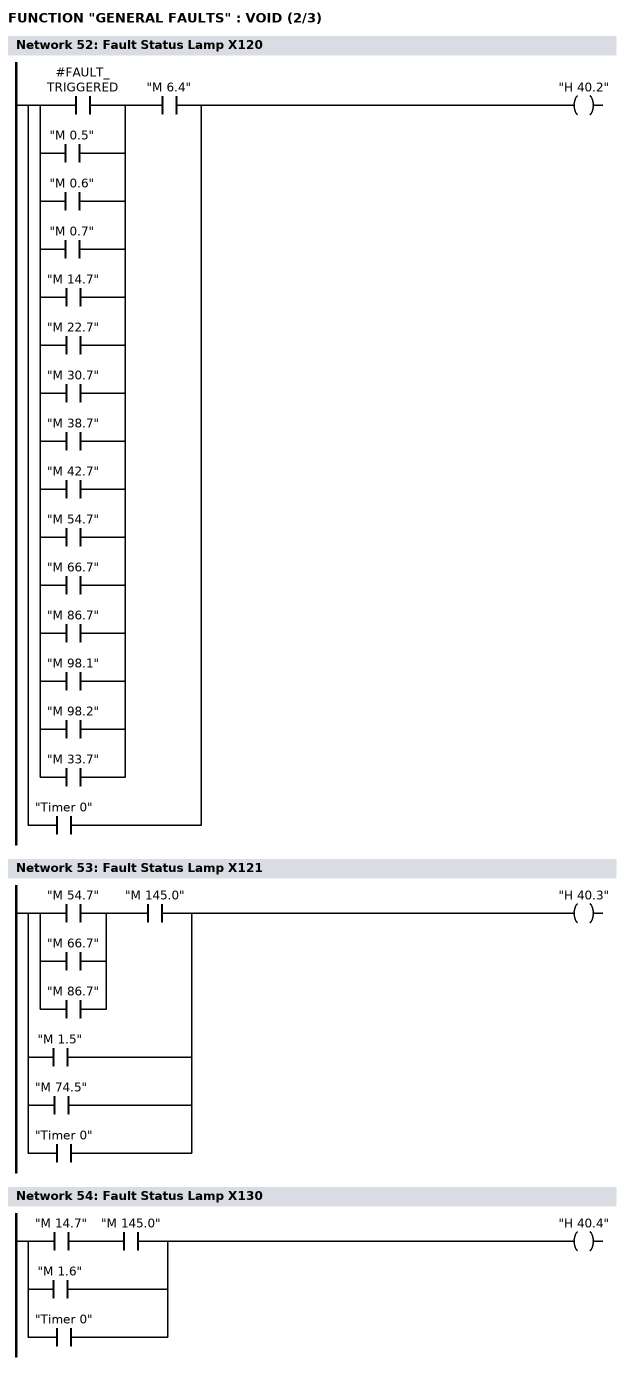

      A(    ;
      O     #FAULT_TRIGGERED;
      O     "M 0.5";
      O     "M 0.6";
      O     "M 0.7";
      O     "M 14.7";
      O     "M 22.7";
      O     "M 30.7";
      O     "M 38.7";
      O     "M 42.7";
      O     "M 54.7";
      O     "M 66.7";
      O     "M 86.7";
      O     "M 98.1";
      O     "M 98.2";
      O     "M 33.7";
      )     ;
      A     "M 6.4";
      O     "Timer 0";
      =     "H 40.2";
NETWORK
TITLE =Fault Status Lamp X121

      A(    ;
      O     "M 54.7";
      O     "M 66.7";
      O     "M 86.7";
      )     ;
      A     "M 145.0";
      O     "M 1.5";
      O     "M 74.5";
      O     "Timer 0";
      =     "H 40.3";
NETWORK
TITLE =Fault Status Lamp X130

      A     "M 14.7";
      A     "M 145.0";
      O     "M 1.6";
      O     "Timer 0";
      =     "H 40.4";
NETWORK
TITLE =Fault Status Lamp X134
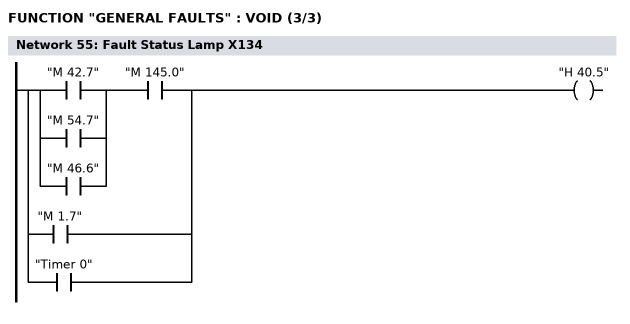

      A(    ;
      O     "M 42.7";
      O     "M 54.7";
      O     "M 46.6";
      )     ;
      A     "M 145.0";
      O     "M 1.7";
      O     "Timer 0";
      =     "H 40.5";
NETWORK
TITLE =Elevator OverTemp

      A     "M 0.6";
      AN    "E 0.3";
      L     W#16#1;
      T     "MB 181";
      BEC   ;
NETWORK
TITLE =Turntable OverTemp

      A     "M 0.6";
      AN    "E 0.4";
      L     W#16#2;
      T     "MB 181";
      BEC   ;
NETWORK
TITLE =Loader OverTemp

      A     "M 0.6";
      AN    "E 0.5";
      L     W#16#3;
      T     "MB 181";
      BEC   ;
NETWORK
TITLE =Conveyor 4 Collator OverTemp

      A     "M 0.6";
      AN    "E 14.0";
      L     W#16#4;
      T     "MB 181";
      BEC   ;
NETWORK
TITLE =Conveyor 6 Delivery OverTemp

      A     "M 0.6";
      AN    "E 14.1";
      L     W#16#5;
      T     "MB 181";
      BEC   ;
NETWORK
TITLE =Pivot Conveyor 10 OverTemp

      A(    ;
      ON    "E 14.2";
      ON    "E 14.3";
      )     ;
      A     "M 0.6";
      O     ;
      A(    ;
      O     "E 14.6";
      O     "E 14.7";
      )     ;
      A     "M 0.6";
      L     W#16#6;
      T     "MB 181";
      BEC   ;
NETWORK
TITLE =OverTemp

      A     "M 0.6";
      A     "E 35.0";
      L     W#16#8;
      T     "MB 181";
      BEC   ;
NETWORK
TITLE =OverTemp

      A     "M 0.6";
      A     "E 35.1";
      L     W#16#9;
      T     "MB 181";
      BEC   ;
NETWORK
TITLE =OverTemp

      A     "M 0.6";
      A     "E 14.6";
      L     W#16#B;
      T     "MB 181";
      BEC   ;
NETWORK
TITLE =OverTemp

      A     "M 0.6";
      A     "E 14.7";
      L     W#16#C;
      T     "MB 181";
      BEC   ;
NETWORK
TITLE =

      A     #FAULT_TRIGGERED;
      A     "M 3.0";
      L     W#16#0;
      T     MB   183;
      BEC   ;
NETWORK
TITLE =

      A     #FAULT_TRIGGERED;
      A     "M 3.1";
      L     W#16#1;
      T     MB   183;
      BEC   ;
NETWORK
TITLE =

      A     #FAULT_TRIGGERED;
      A     "M 3.2";
      L     W#16#2;
      T     MB   183;
      BEC   ;
NETWORK
TITLE =

      A     #FAULT_TRIGGERED;
      A     "M 3.3";
      L     W#16#3;
      T     MB   183;
      BEC   ;
NETWORK
TITLE =

      A     #FAULT_TRIGGERED;
      A     "M 3.4";
      L     W#16#4;
      T     MB   183;
      BEC   ;
NETWORK
TITLE =

      A     #FAULT_TRIGGERED;
      A     "M 3.5";
      L     W#16#5;
      T     MB   183;
      BEC   ;
NETWORK
TITLE =

      A     #FAULT_TRIGGERED;
      A     "M 3.6";
      L     W#16#6;
      T     MB   183;
      BEC   ;
NETWORK
TITLE =

      A     #FAULT_TRIGGERED;
      A     "M 3.7";
      L     W#16#7;
      T     MB   183;
      BEC   ;
NETWORK
TITLE =

      A     #FAULT_TRIGGERED;
      A     "M 4.0";
      L     W#16#8;
      T     MB   182;
      BEC   ;
NETWORK
TITLE =

      A     #FAULT_TRIGGERED;
      A     "M 4.1";
      L     W#16#9;
      T     MB   182;
      BEC   ;
NETWORK
TITLE =

      A     #FAULT_TRIGGERED;
      A     "M 4.2";
      L     W#16#10;
      T     MB   182;
      BEC   ;
NETWORK
TITLE =

      A     #FAULT_TRIGGERED;
      A     "M 4.3";
      L     W#16#11;
      T     MB   182;
      BEC   ;
NETWORK
TITLE =

      A     #FAULT_TRIGGERED;
      A     "M 4.4";
      L     W#16#12;
      T     MB   182;
      BEC   ;
NETWORK
TITLE =

      A     #FAULT_TRIGGERED;
      A     "M 4.5";
      L     W#16#13;
      T     MB   182;
      BEC   ;
NETWORK
TITLE =

      A     #FAULT_TRIGGERED;
      A     "M 4.6";
      L     W#16#14;
      T     MB   182;
      BEC   ;
NETWORK
TITLE =

      L     W#16#0;
      T     "MW 180";
      T     MW   182;
END_FUNCTION

FUNCTION "BLINKER" : VOID
TITLE =Blinker
VERSION : 0.0

BEGIN
NETWORK
TITLE =
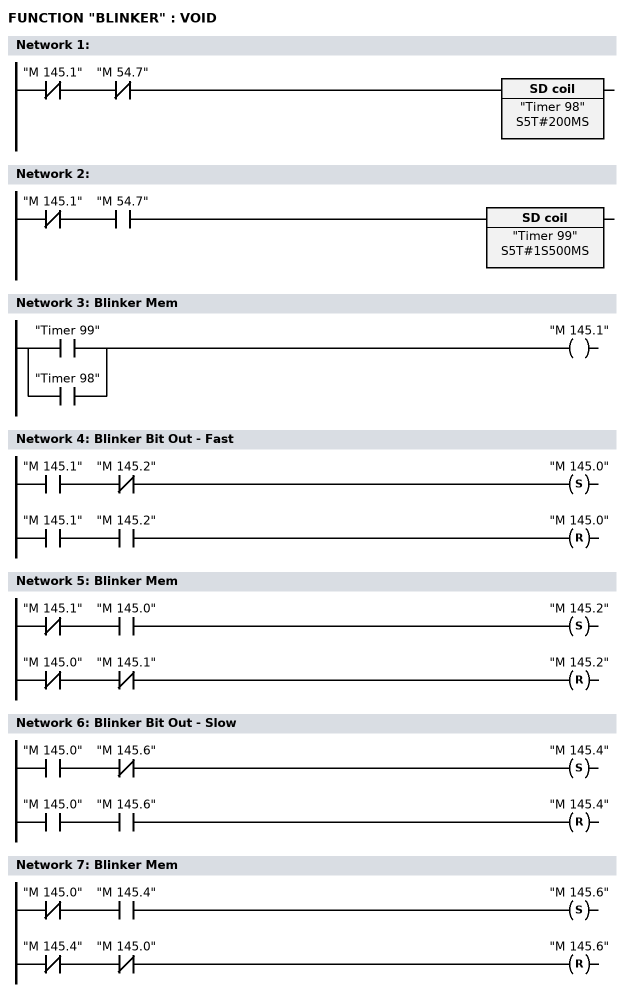

      AN    "M 145.1";
      AN    "M 54.7";
      L     S5T#200MS;
      SD    "Timer 98";
NETWORK
TITLE =

      AN    "M 145.1";
      A     "M 54.7";
      L     S5T#1S500MS;
      SD    "Timer 99";
NETWORK
TITLE =Blinker Mem

      O     "Timer 99";
      O     "Timer 98";
      =     "M 145.1";
NETWORK
TITLE =Blinker Bit Out - Fast

      A     "M 145.1";
      AN    "M 145.2";
      S     "M 145.0";
//;
      A     "M 145.1";
      A     "M 145.2";
      R     "M 145.0";
NETWORK
TITLE =Blinker Mem

      AN    "M 145.1";
      A     "M 145.0";
      S     "M 145.2";
//;
      AN    "M 145.0";
      AN    "M 145.1";
      R     "M 145.2";
NETWORK
TITLE =Blinker Bit Out - Slow

      A     "M 145.0";
      AN    "M 145.6";
      S     "M 145.4";
//;
      A     "M 145.0";
      A     "M 145.6";
      R     "M 145.4";
NETWORK
TITLE =Blinker Mem

      AN    "M 145.0";
      A     "M 145.4";
      S     "M 145.6";
//;
      AN    "M 145.4";
      AN    "M 145.0";
      R     "M 145.6";
END_FUNCTION

FUNCTION "LIGHT CURTAIN - SAFETY" : VOID
TITLE =Conveyors Catways - Access Safety
//Access to Conveyor 1-2-3 & 4 : Crossing Light Curtains Latches / Freezes these
//Conveyors !
//- To Resume Run, CatWay 1 (Conveyors 1-2-3) :  Push Top PB (Catway)
//and Push Lower PB (Main Floor) within 15sec .
//- To Resume Run, CatWay 2 (Conveyors 3-4) :  Push Top PB (Catway) .
//
//If Crossing CatWay 2 Light Curtain while No Conveyors are running, Run will
//resume automatic after 1 sec of free Light Curtain.
//
//Big Red Light will Blink to confirm the Conveyors are disabled / Safe .
VERSION : 0.1

BEGIN
NETWORK
TITLE =Safety Light Curtains -  Trigger 2 - Momentary SF = 1s
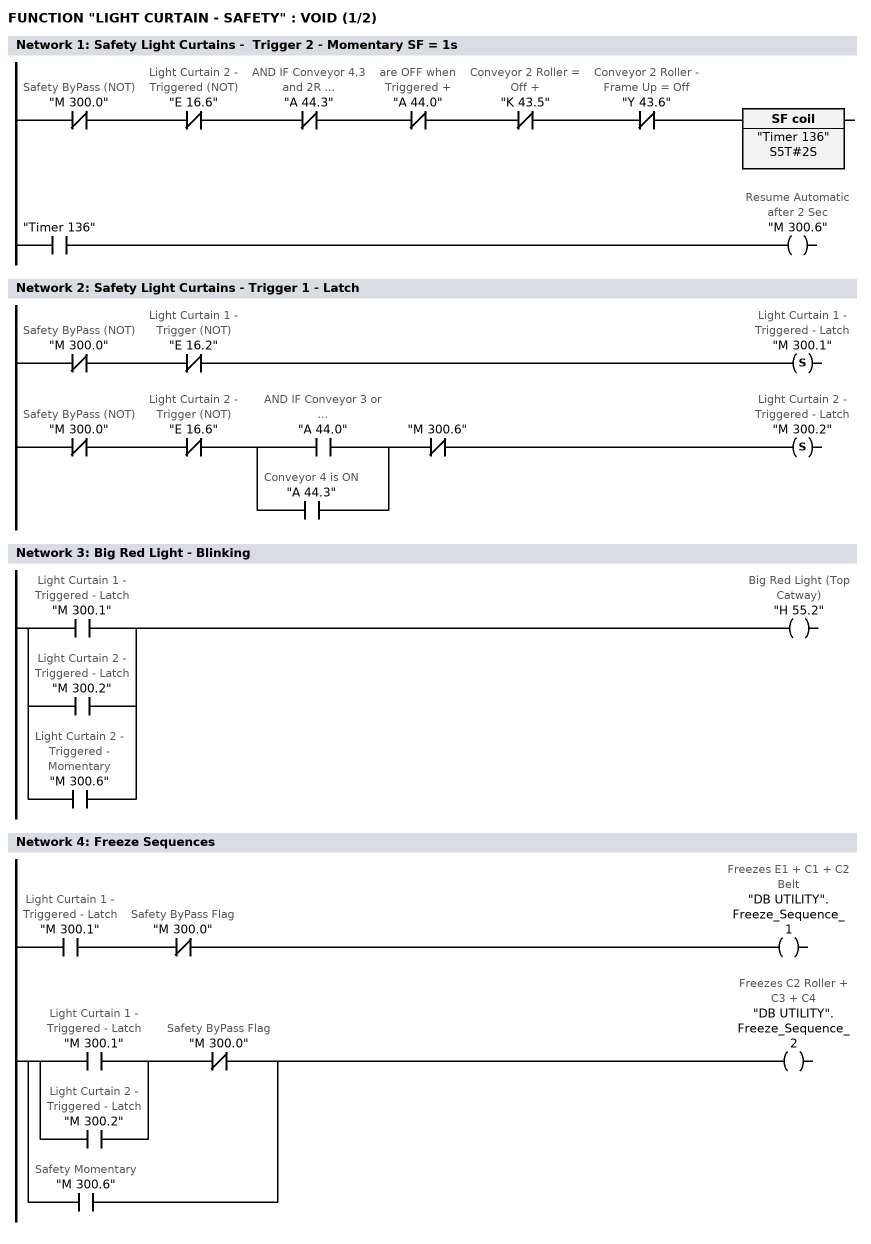

      AN    "M 300.0"; // Safety ByPass (NOT)
      AN    "E 16.6"; // Light Curtain 2 - Triggered (NOT)
      AN    "A 44.3"; // AND IF Conveyor 4,3 and 2R ...
      AN    "A 44.0"; // are OFF when Triggered +
      AN    "K 43.5"; // Conveyor 2 Roller = Off +
      AN    "Y 43.6"; // Conveyor 2 Roller - Frame Up = Off
      L     S5T#2S;
      SF    "Timer 136"; // Debouncer 2s
//;
      A     "Timer 136";
      =     "M 300.6"; // Resume Automatic after 2 Sec

NETWORK
TITLE =Safety Light Curtains - Trigger 1 - Latch

      AN    "M 300.0"; // Safety ByPass (NOT)
      AN    "E 16.2"; // Light Curtain 1 - Trigger (NOT)
      S     "M 300.1"; // Light Curtain 1 - Triggered - Latch
//;
      AN    "M 300.0"; // Safety ByPass (NOT)
      AN    "E 16.6"; // Light Curtain 2 - Trigger (NOT)
      A(    ;
      O     "A 44.0"; // AND IF Conveyor 3 or ...
      O     "A 44.3"; // Conveyor 4 is ON
      )     ;
      AN    "M 300.6";
      S     "M 300.2"; // Light Curtain 2 - Triggered - Latch
NETWORK
TITLE =Big Red Light - Blinking

      A(    ;
      O     "M 300.1"; // Light Curtain 1 - Triggered - Latch
      O     "M 300.2"; // Light Curtain 2 - Triggered - Latch
      O     "M 300.6"; // Light Curtain 2 - Triggered - Momentary
      )     ;
      =     "H 55.2"; // Big Red Light (Top Catway)
NETWORK
TITLE =Freeze Sequences

      A     "M 300.1"; // Light Curtain 1 - Triggered - Latch
      AN    "M 300.0"; // Safety ByPass Flag
      =     "DB UTILITY".Freeze_Sequence_1; //   Freezes E1 + C1 + C2 Belt
//;
      A     "M 300.1"; // Light Curtain 1 - Triggered - Latch
      O     "M 300.2"; // Light Curtain 2 - Triggered - Latch
      AN    "M 300.0"; // Safety ByPass Flag
      O     "M 300.6"; // Safety Momentary
      =     "DB UTILITY".Freeze_Sequence_2; //  Freezes C2 Roller + C3 + C4
NETWORK
TITLE =Safety ByPass - While blocking Curtain, Push Top Button for 5s
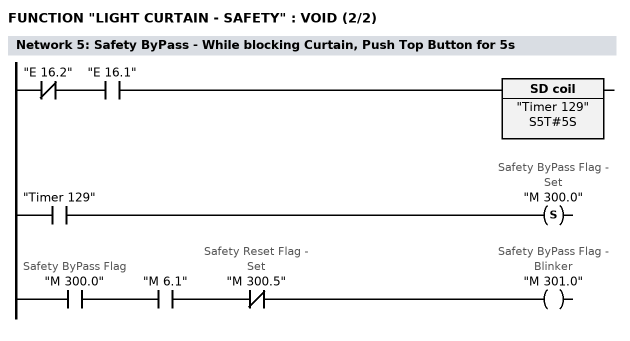

      AN    "E 16.2";
      A     "E 16.1";
      L     S5T#5S;
      SD    "Timer 129";
//;
      A     "Timer 129";
      S     "M 300.0"; // Safety ByPass Flag - Set
//;
      A     "M 300.0"; // Safety ByPass Flag
      A     "M 6.1";
      AN    "M 300.5"; // Safety Reset Flag - Set
      =     "M 301.0"; // Safety ByPass Flag - Blinker

NETWORK
TITLE =TEST REMOTE B+

      R     "A 58.4";

NETWORK
TITLE =PB Led - Control
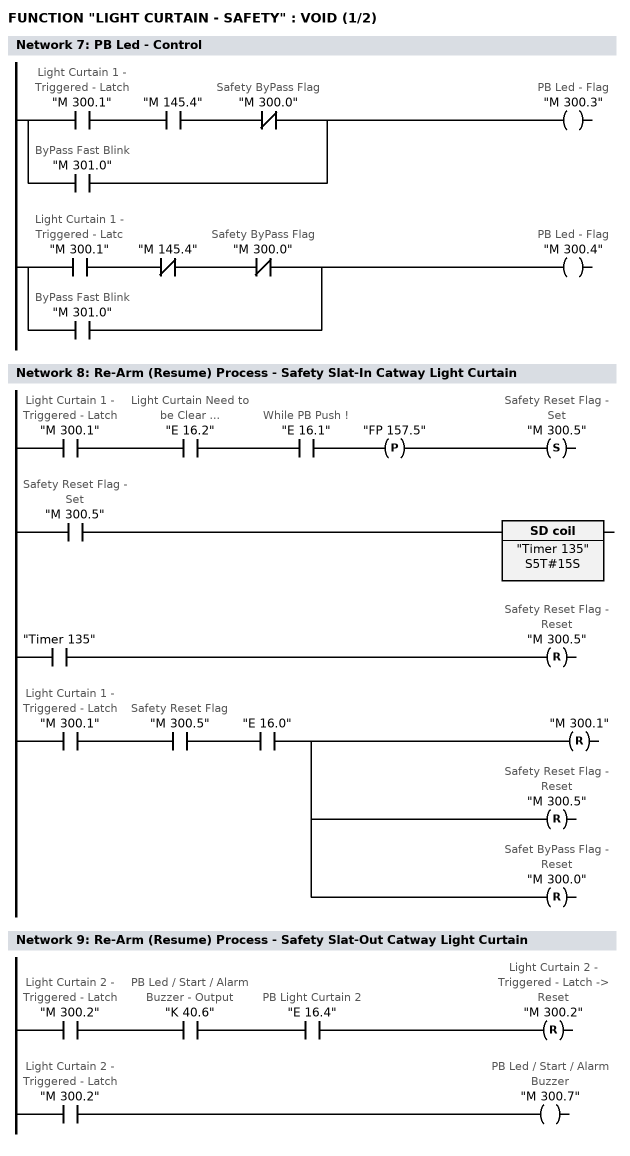

      A     "M 300.1"; // Light Curtain 1 - Triggered - Latch
      A     "M 145.4";
      AN    "M 300.0"; // Safety ByPass Flag
      O     "M 301.0"; // ByPass Fast Blink
      =     "M 300.3"; // PB Led - Flag
//;
      A     "M 300.1"; // Light Curtain 1 - Triggered - Latc
      AN    "M 145.4";
      AN    "M 300.0"; // Safety ByPass Flag
      O     "M 301.0"; // ByPass Fast Blink
      =     "M 300.4"; // PB Led - Flag
NETWORK
TITLE =Re-Arm (Resume) Process - Safety Slat-In Catway Light Curtain

      A     "M 300.1"; // Light Curtain 1 - Triggered - Latch
      A     "E 16.2"; // Light Curtain Need to be Clear ...
      A     "E 16.1"; // While PB Push !
      FP    "FP 157.5";
      S     "M 300.5"; // Safety Reset Flag - Set
//;
      A     "M 300.5"; // Safety Reset Flag - Set
      L     S5T#15S;
      SD    "Timer 135"; // Safety Reset Flag - TimeOut
//;
      A     "Timer 135";
      R     "M 300.5"; // Safety Reset Flag - Reset
//;
      A     "M 300.1"; // Light Curtain 1 - Triggered - Latch
      A     "M 300.5"; // Safety Reset Flag
      A     "E 16.0";
      R     "M 300.1";
      R     "M 300.5"; // Safety Reset Flag - Reset
      R     "M 300.0"; // Safet ByPass Flag - Reset
NETWORK
TITLE =Re-Arm (Resume) Process - Safety Slat-Out Catway Light Curtain

      A     "M 300.2"; // Light Curtain 2 - Triggered - Latch
      A     "K 40.6"; // PB Led / Start / Alarm Buzzer - Output
      A     "E 16.4"; // PB Light Curtain 2
      R     "M 300.2"; // Light Curtain 2 - Triggered - Latch -> Reset
//;
      A     "M 300.2"; // Light Curtain 2 - Triggered - Latch
      =     "M 300.7"; // PB Led / Start / Alarm Buzzer
NETWORK
TITLE =PB Led - Out
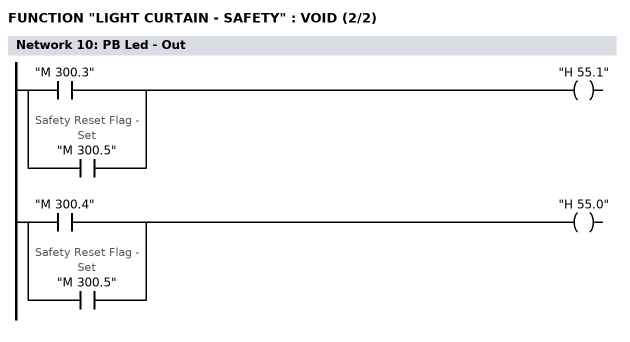

      A     "M 300.3";
      O     "M 300.5"; // Safety Reset Flag - Set
      =     "H 55.1";
//;
      A     "M 300.4";
      O     "M 300.5"; // Safety Reset Flag - Set
      =     "H 55.0";
END_FUNCTION

FUNCTION "CONVEYORS CLEARING" : VOID
TITLE =Conveyors - Clearing Function
//New Order Sequence
NAME : CLEARING
VERSION : 0.0


VAR_TEMP
  EMPTY_11 : BOOL ;	//Empty Conveyor 11
  EMPTY_21 : BOOL ;	//Empty Conveyor 21
  EMPTY_12_22 : BOOL ;	//Empty Conveyor 12 & 22
  EMPTY_13_23 : BOOL ;	//Empty Conveyor 13 & 23
  C10_EMPTY_TEST : BOOL ;
  CLEARING_ABORT : BOOL ;
END_VAR
BEGIN
NETWORK
TITLE =HMI Clearing Call

      A     "M 140.3";
      A     "HMI_DB".CLEARING_SSW_MAIN;
      =     "M 5.2";
//;
      L     8;
      A     "M 10.0";
      =     "HMI_DB".CLEARING_SSW_STATUS;
      JC    CLEA;
      L     0;

CLEA: T     "HMI_DB".CLEARING_FUNCTION;

      A     "M 10.0";
      FN    "FN 155.7";
      R     "HMI_DB".CLEARING_SSW_MAIN;
      R     "M 54.2";
//;
      A     "M 5.2";
      FP    "FP 147.4";
      AN    "B 10.7"; // C11 - Empty
      AN    "B 11.0"; // C12 - Empty
      AN    "B 11.1"; // C13 - Empty
      AN    "B 11.2"; // C13 - Empty
      AN    "B 15.4"; // C21 - Empty
      AN    "B 15.5"; // C22 - Empty
      AN    "B 15.6"; // C23 - Empty
      AN    "B 15.7"; // C23 - Empty
      S     "M 54.2"; // Empty C11...C23
NETWORK
TITLE =New Order Seq - First New Order Packet to Pivot Conveyor 10
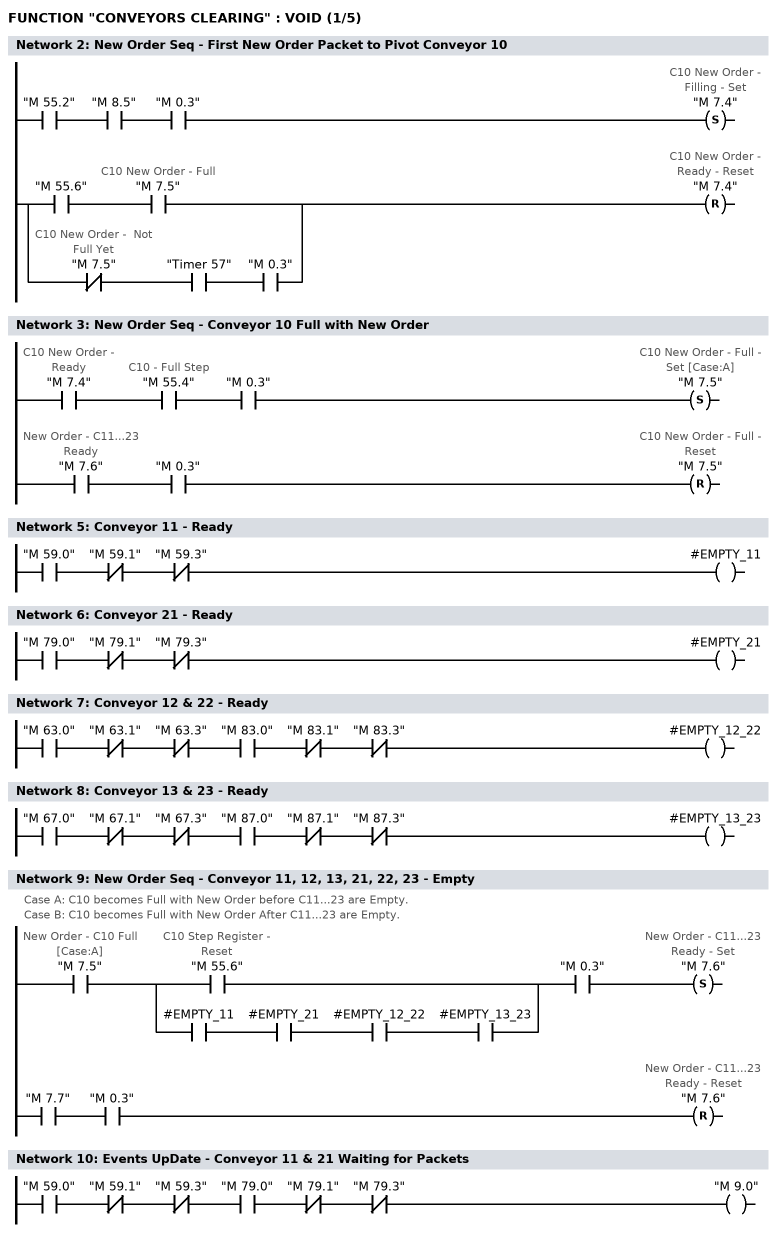

      A     "M 55.2";
      A     "M 8.5";
      A     "M 0.3";
      S     "M 7.4"; // C10 New Order - Filling - Set
//;
      A(    ;
      A     "M 55.6";
      A     "M 7.5"; // C10 New Order - Full
      O     ;
      AN    "M 7.5"; // C10 New Order -  Not Full Yet
      A     "Timer 57";
      A     "M 0.3";
      )     ;
      R     "M 7.4"; // C10 New Order - Ready - Reset
NETWORK
TITLE =New Order Seq - Conveyor 10 Full with New Order

      A     "M 7.4"; // C10 New Order - Ready
      A     "M 55.4"; // C10 - Full Step
      A     "M 0.3";
      S     "M 7.5"; // C10 New Order - Full - Set [Case:A]
//;
      A     "M 7.6"; // New Order - C11...23 Ready
      A     "M 0.3";
      R     "M 7.5"; // C10 New Order - Full - Reset
NETWORK
TITLE =New Order Seq
//New Order Seq - Waiting for the last Order Packets to Run out !


NETWORK
TITLE =Conveyor 11 - Ready

      A     "M 59.0";
      AN    "M 59.1";
      AN    "M 59.3";
      =     #EMPTY_11;
NETWORK
TITLE =Conveyor 21 - Ready

      A     "M 79.0";
      AN    "M 79.1";
      AN    "M 79.3";
      =     #EMPTY_21;
NETWORK
TITLE =Conveyor 12 & 22 - Ready

      A     "M 63.0";
      AN    "M 63.1";
      AN    "M 63.3";
      A     "M 83.0";
      AN    "M 83.1";
      AN    "M 83.3";
      =     #EMPTY_12_22;
NETWORK
TITLE =Conveyor 13 & 23 - Ready

      A     "M 67.0";
      AN    "M 67.1";
      AN    "M 67.3";
      A     "M 87.0";
      AN    "M 87.1";
      AN    "M 87.3";
      =     #EMPTY_13_23;
NETWORK
TITLE =New Order Seq - Conveyor 11, 12, 13, 21, 22, 23 - Empty
//Case A: C10 becomes Full with New Order before C11...23 are Empty.
//Case B: C10 becomes Full with New Order After C11...23 are Empty.
      A     "M 7.5"; // New Order - C10 Full [Case:A]
      A(    ;
      A     "M 55.6"; // C10 Step Register - Reset
      O     ;
      A     #EMPTY_11;
      A     #EMPTY_21;
      A     #EMPTY_12_22;
      A     #EMPTY_13_23;
      )     ;
      A     "M 0.3";
      S     "M 7.6"; // New Order - C11...23 Ready - Set
//;
      A     "M 7.7";
      A     "M 0.3";
      R     "M 7.6"; // New Order - C11...23 Ready - Reset
NETWORK
TITLE =Events UpDate - Conveyor 11 & 21 Waiting for Packets

      A     "M 59.0";
      AN    "M 59.1";
      AN    "M 59.3";
      A     "M 79.0";
      AN    "M 79.1";
      AN    "M 79.3";
      =     "M 9.0";
NETWORK
TITLE =New Order Seq - Conveyors 11, 21 - Empty
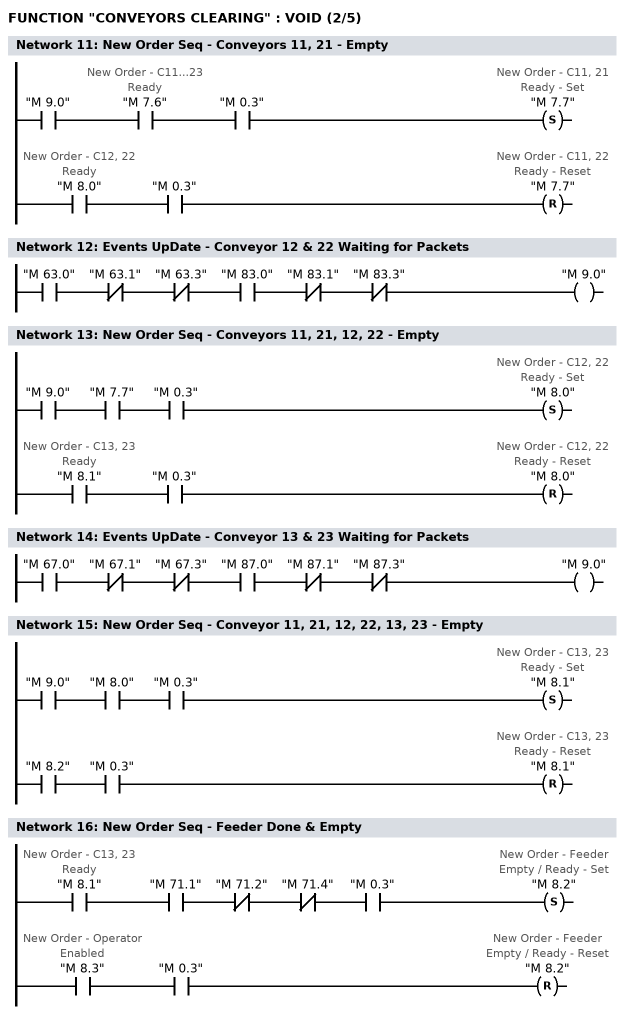

      A     "M 9.0";
      A     "M 7.6"; // New Order - C11...23 Ready
      A     "M 0.3";
      S     "M 7.7"; // New Order - C11, 21 Ready - Set
//;
      A     "M 8.0"; // New Order - C12, 22 Ready
      A     "M 0.3";
      R     "M 7.7"; // New Order - C11, 22 Ready - Reset
NETWORK
TITLE =Events UpDate - Conveyor 12 & 22 Waiting for Packets

      A     "M 63.0";
      AN    "M 63.1";
      AN    "M 63.3";
      A     "M 83.0";
      AN    "M 83.1";
      AN    "M 83.3";
      =     "M 9.0";
NETWORK
TITLE =New Order Seq - Conveyors 11, 21, 12, 22 - Empty

      A     "M 9.0";
      A     "M 7.7";
      A     "M 0.3";
      S     "M 8.0"; // New Order - C12, 22 Ready - Set
//;
      A     "M 8.1"; // New Order - C13, 23 Ready
      A     "M 0.3";
      R     "M 8.0"; // New Order - C12, 22 Ready - Reset
NETWORK
TITLE =Events UpDate - Conveyor 13 & 23 Waiting for Packets

      A     "M 67.0";
      AN    "M 67.1";
      AN    "M 67.3";
      A     "M 87.0";
      AN    "M 87.1";
      AN    "M 87.3";
      =     "M 9.0";
NETWORK
TITLE =New Order Seq - Conveyor 11, 21, 12, 22, 13, 23 - Empty

      A     "M 9.0";
      A     "M 8.0";
      A     "M 0.3";
      S     "M 8.1"; // New Order - C13, 23 Ready - Set
//;
      A     "M 8.2";
      A     "M 0.3";
      R     "M 8.1"; // New Order - C13, 23 Ready - Reset
NETWORK
TITLE =New Order Seq - Feeder Done & Empty

      A     "M 8.1"; // New Order - C13, 23 Ready
      A     "M 71.1";
      AN    "M 71.2";
      AN    "M 71.4";
      A     "M 0.3";
      S     "M 8.2"; // New Order - Feeder Empty / Ready - Set
//;
      A     "M 8.3"; // New Order - Operator Enabled
      A     "M 0.3";
      R     "M 8.2"; // New Order - Feeder Empty / Ready - Reset
NETWORK
TITLE =Conveyor 10 Clearing Enable after New Order
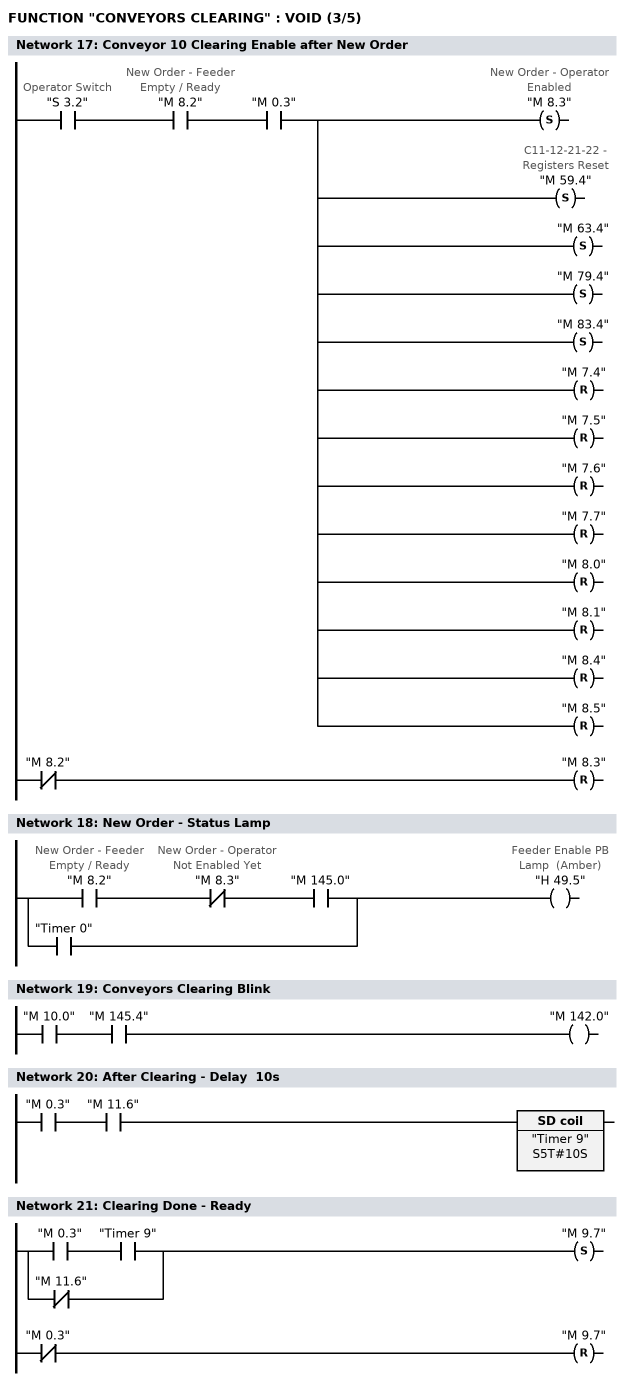

      A     "S 3.2"; // Operator Switch
      A     "M 8.2"; // New Order - Feeder Empty / Ready
      A     "M 0.3";
      S     "M 8.3"; // New Order - Operator Enabled
      S     "M 59.4"; // C11-12-21-22 - Registers Reset
      S     "M 63.4";
      S     "M 79.4";
      S     "M 83.4";
//;
      R     "M 7.4";
      R     "M 7.5";
      R     "M 7.6";
      R     "M 7.7";
      R     "M 8.0";
      R     "M 8.1";
      R     "M 8.4";
      R     "M 8.5";
//;
      ON    "M 8.2";
      R     "M 8.3";
NETWORK
TITLE =New Order - Status Lamp

      A     "M 8.2"; // New Order - Feeder Empty / Ready
      AN    "M 8.3"; // New Order - Operator Not Enabled Yet
      A     "M 145.0";
      O     "Timer 0";
      =     "H 49.5"; // Feeder Enable PB Lamp  (Amber)
NETWORK
TITLE =Conveyors Clearing Blink

      A     "M 10.0";
      A     "M 145.4";
      =     "M 142.0";
NETWORK
TITLE =After Clearing - Delay  10s

      A     "M 0.3";
      A     "M 11.6";
      L     S5T#10S;
      SD    "Timer 9";
NETWORK
TITLE =Clearing Done - Ready

      A     "M 0.3";
      A     "Timer 9";
      ON    "M 11.6";
      S     "M 9.7";
//;
      ON    "M 0.3";
      R     "M 9.7";
NETWORK
TITLE =Clearing Command
//Clearing Command


NETWORK
TITLE =Conveyors Clearing - Cmd
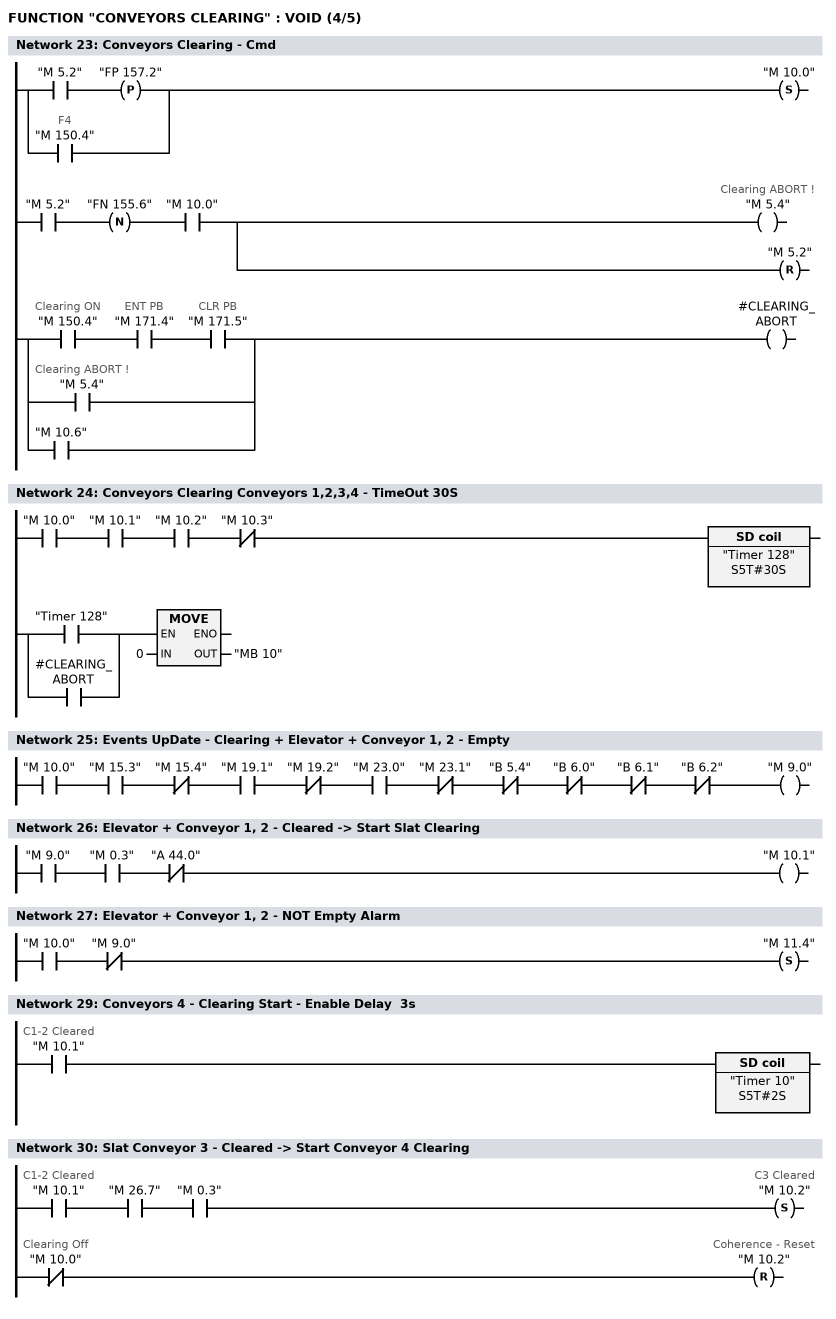

      A(    ;
      A     "M 5.2";
      FP    "FP 157.2";
      O     ;
      A     "M 150.4"; // F4
      )     ;
      S     "M 10.0";
//;
      A     "M 5.2";
      FN    "FN 155.6";
      A     "M 10.0";
      =     "M 5.4"; // Clearing ABORT !
      R     "M 5.2";
//;
      A(    ;
      A     "M 150.4"; // Clearing ON
      A     "M 171.4"; // ENT PB
      A     "M 171.5"; // CLR PB
      O     "M 5.4"; // Clearing ABORT !
      O     "M 10.6";
      )     ;
      =     #CLEARING_ABORT;
NETWORK
TITLE =Conveyors Clearing Conveyors 1,2,3,4 - TimeOut 30S

      A     "M 10.0";
      A     "M 10.1";
      A     "M 10.2";
      AN    "M 10.3";
      L     S5T#30S;
      SD    "Timer 128";
//;
      A     "Timer 128";
      O     #CLEARING_ABORT;
      JNB   NCLR;
      L     0;
      T     "MB 10"; // Clearing OFF

NCLR: NOP   0;
NETWORK
TITLE =Events UpDate - Clearing + Elevator + Conveyor 1, 2 - Empty

      A     "M 10.0";
      A     "M 15.3";
      AN    "M 15.4";
      A     "M 19.1";
      AN    "M 19.2";
      A     "M 23.0";
      AN    "M 23.1";
      AN    "B 5.4";
      AN    "B 6.0";
      AN    "B 6.1";
      AN    "B 6.2";
      =     "M 9.0";
NETWORK
TITLE =Elevator + Conveyor 1, 2 - Cleared -> Start Slat Clearing

      A     "M 9.0";
      A     "M 0.3";
      AN    "A 44.0";
      =     "M 10.1";
NETWORK
TITLE =Elevator + Conveyor 1, 2 - NOT Empty Alarm

      A     "M 10.0";
      AN    "M 9.0";
      S     "M 11.4";
NETWORK
TITLE =Clearing Sequence
//Clearing Sequence from Slat 3 to Pivot 10 Conveyors


NETWORK
TITLE =Conveyors 4 - Clearing Start - Enable Delay  3s

      A     "M 10.1"; // C1-2 Cleared
      L     S5T#2S;
      SD    "Timer 10";
NETWORK
TITLE =Slat Conveyor 3 - Cleared -> Start Conveyor 4 Clearing

      A     "M 10.1"; // C1-2 Cleared
      A     "M 26.7";
      A     "M 0.3";
      S     "M 10.2"; // C3 Cleared
//;
      AN    "M 10.0"; // Clearing Off
      R     "M 10.2"; // Coherence - Reset
NETWORK
TITLE =Conveyors 3, 4 - Cleared -> Start Conveyor 5, 6 Clearing
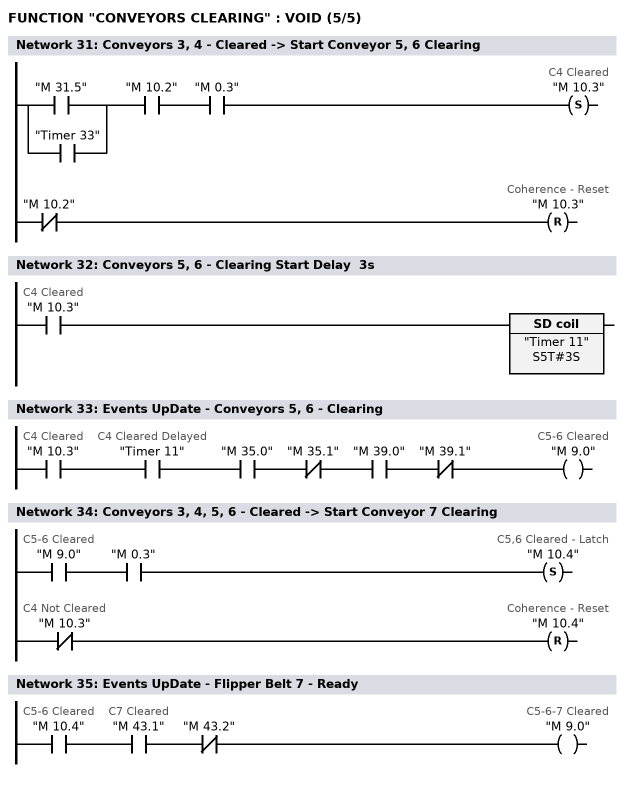

      A(    ;
      O     "M 31.5";
      O     "Timer 33";
      )     ;
      A     "M 10.2";
      A     "M 0.3";
      S     "M 10.3"; // C4 Cleared
//;
      AN    "M 10.2";
      R     "M 10.3"; // Coherence - Reset
NETWORK
TITLE =Conveyors 5, 6 - Clearing Start Delay  3s

      A     "M 10.3"; // C4 Cleared
      L     S5T#3S;
      SD    "Timer 11"; // C4 Cleared Delayed
NETWORK
TITLE =Events UpDate - Conveyors 5, 6 - Clearing

      A     "M 10.3"; // C4 Cleared
      A     "Timer 11"; // C4 Cleared Delayed
      A     "M 35.0";
      AN    "M 35.1";
      A     "M 39.0";
      AN    "M 39.1";
      =     "M 9.0"; // C5-6 Cleared
NETWORK
TITLE =Conveyors 3, 4, 5, 6 - Cleared -> Start Conveyor 7 Clearing

      A     "M 9.0"; // C5-6 Cleared
      A     "M 0.3";
      S     "M 10.4"; // C5,6 Cleared - Latch
//;
      AN    "M 10.3"; // C4 Not Cleared
      R     "M 10.4"; // Coherence - Reset
NETWORK
TITLE =Events UpDate - Flipper Belt 7 - Ready

      A     "M 10.4"; // C5-6 Cleared
      A     "M 43.1"; // C7 Cleared
      AN    "M 43.2";
      =     "M 9.0"; // C5-6-7 Cleared
NETWORK
TITLE =Conveyors 3, 4, 5, 6, 7, 8, 9 - Clearing - Cleared / Ready

      A     "M 9.0"; // C5-6-7 Cleared
      A     "M 47.2"; // C8 Cleared
      AN    "M 47.3";
      A     "M 51.1"; // C9 Cleared
      AN    "M 51.2";
      AN    "B 9.7"; // C9 - Pusher2 - Edge Cleared
      A     "M 0.3";
      L     S5T#3S;
      SD    "Timer 56"; // Delay 3s
//;
      A     "Timer 56";
      =     "M 10.5"; // C10 UpStream Cleared
      FP    "M 188.4";
      S     "M 58.2"; // C10 UpStream Cleared - Trigger Set
//;
      A     "M 10.5";
      L     S5T#1S;
      SE    "Timer 58"; // UpStream Cleared - Pulse 1s
NETWORK
TITLE =Pivot Conveyor 10 - Clearing - Cleared / Ready
//"C10_EMPTY_TEST" : Work Around to "Will NOT Empty Conveyor 10 - Pivot after a
//Clearing (F4)".
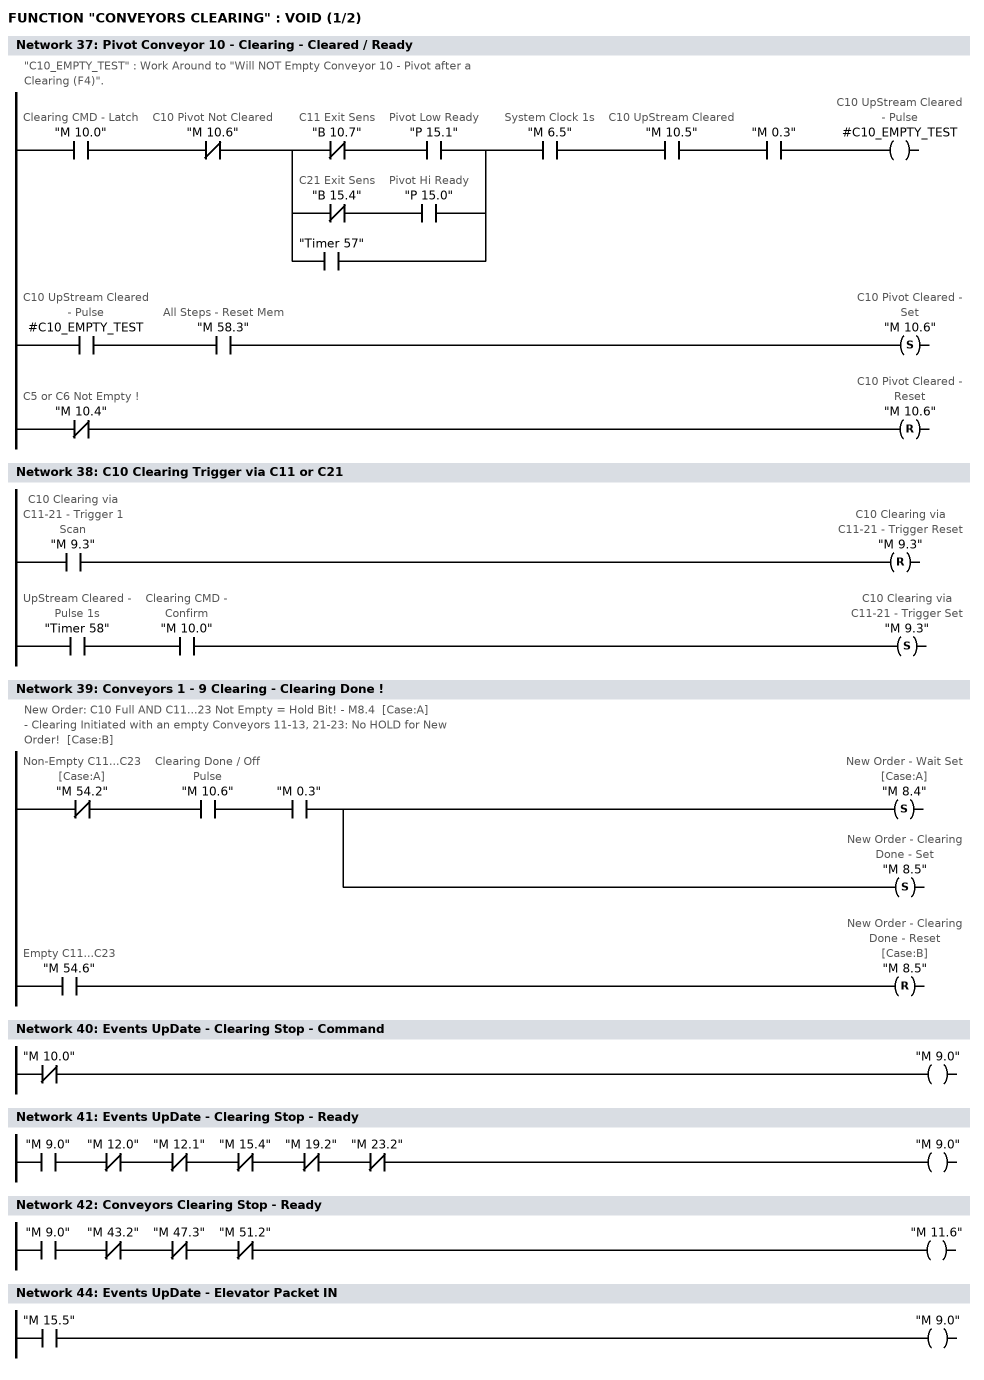
      A     "M 10.0"; // Clearing CMD - Latch
      AN    "M 10.6"; // C10 Pivot Not Cleared
      A(    ;
      AN    "B 10.7"; // C11 Exit Sens
      A     "P 15.1"; // Pivot Low Ready
      O     ;
      AN    "B 15.4"; // C21 Exit Sens
      A     "P 15.0"; // Pivot Hi Ready
      O     "Timer 57";
      )     ;
      A     "M 6.5"; // System Clock 1s
      A     "M 10.5"; // C10 UpStream Cleared
      A     "M 0.3";
      =     #C10_EMPTY_TEST; // C10 UpStream Cleared - Pulse
//;
      A     #C10_EMPTY_TEST; // C10 UpStream Cleared - Pulse
      A     "M 58.3"; // All Steps - Reset Mem
      S     "M 10.6"; // C10 Pivot Cleared - Set
//;
      AN    "M 10.4"; // C5 or C6 Not Empty !
      R     "M 10.6"; // C10 Pivot Cleared - Reset
NETWORK
TITLE =C10 Clearing Trigger via C11 or C21

      A     "M 9.3"; // C10 Clearing via C11-21 - Trigger 1 Scan
      R     "M 9.3"; // C10 Clearing via C11-21 - Trigger Reset
//;
      A     "Timer 58"; // UpStream Cleared - Pulse 1s
      A     "M 10.0"; // Clearing CMD - Confirm
      S     "M 9.3"; // C10 Clearing via C11-21 - Trigger Set
NETWORK
TITLE =Conveyors 1 - 9 Clearing - Clearing Done !
//New Order: C10 Full AND C11...23 Not Empty = Hold Bit! - M8.4  [Case:A]
//
//- Clearing Initiated with an empty Conveyors 11-13, 21-23: No HOLD for New
//Order!  [Case:B]
//
      AN    "M 54.2"; // Non-Empty C11...C23   [Case:A]
      A     "M 10.6"; // Clearing Done / Off Pulse
      A     "M 0.3";
      S     "M 8.4"; // New Order - Wait Set   [Case:A]
      S     "M 8.5"; // New Order - Clearing Done - Set
//;
      A     "M 54.6"; // Empty C11...C23
      R     "M 8.5"; // New Order - Clearing Done - Reset   [Case:B]
NETWORK
TITLE =Events UpDate - Clearing Stop - Command

      AN    "M 10.0";
      =     "M 9.0";
NETWORK
TITLE =Events UpDate - Clearing Stop - Ready

      A     "M 9.0";
      AN    "M 12.0";
      AN    "M 12.1";
      AN    "M 15.4";
      AN    "M 19.2";
      AN    "M 23.2";
      =     "M 9.0";
NETWORK
TITLE =Conveyors Clearing Stop - Ready

      A     "M 9.0";
      AN    "M 43.2";
      AN    "M 47.3";
      AN    "M 51.2";
      =     "M 11.6";
NETWORK
TITLE =New Order
//New Order : Start Filling Conveyors


NETWORK
TITLE =Events UpDate - Elevator Packet IN

      A     "M 15.5";
      =     "M 9.0";
NETWORK
TITLE =Events UpDate - Conveyor 1 - 9 - Packet Present
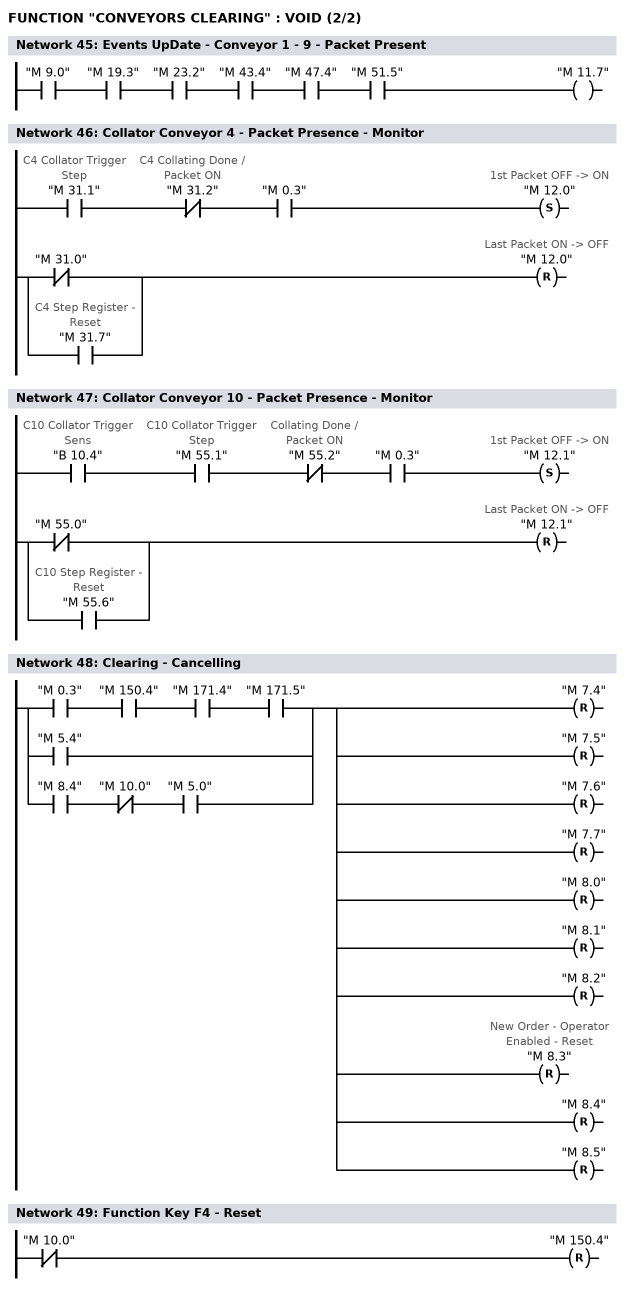

      A     "M 9.0";
      A     "M 19.3";
      A     "M 23.2";
      A     "M 43.4";
      A     "M 47.4";
      A     "M 51.5";
      =     "M 11.7";
NETWORK
TITLE =Collator Conveyor 4 - Packet Presence - Monitor

      A     "M 31.1"; // C4 Collator Trigger Step
      AN    "M 31.2"; // C4 Collating Done / Packet ON
      A     "M 0.3";
      S     "M 12.0"; // 1st Packet OFF -> ON
//;
      A(    ;
      ON    "M 31.0";
      O     "M 31.7"; // C4 Step Register - Reset
      )     ;
      R     "M 12.0"; // Last Packet ON -> OFF
NETWORK
TITLE =Collator Conveyor 10 - Packet Presence - Monitor

      A     "B 10.4"; // C10 Collator Trigger Sens
      A     "M 55.1"; // C10 Collator Trigger Step
      AN    "M 55.2"; // Collating Done / Packet ON
      A     "M 0.3";
      S     "M 12.1"; // 1st Packet OFF -> ON
//;
      A(    ;
      ON    "M 55.0";
      O     "M 55.6"; // C10 Step Register - Reset
      )     ;
      R     "M 12.1"; // Last Packet ON -> OFF
NETWORK
TITLE =Clearing - Cancelling

      A     "M 0.3";
      A     "M 150.4";
      A     "M 171.4";
      A     "M 171.5";
      O     "M 5.4";
      O(    ;
      A     "M 8.4";
      AN    "M 10.0";
      A     "M 5.0";
      )     ;
      R     "M 7.4";
      R     "M 7.5";
      R     "M 7.6";
      R     "M 7.7";
      R     "M 8.0";
      R     "M 8.1";
      R     "M 8.2";
      R     "M 8.3"; // New Order - Operator Enabled - Reset
      R     "M 8.4";
      R     "M 8.5";
NETWORK
TITLE =Function Key F4 - Reset

      AN    "M 10.0";
      R     "M 150.4";
END_FUNCTION

FUNCTION "CONVEYOR 0 + PUSHER 0" : VOID
TITLE =Conveyor 0 & Pusher 0
NAME : 'Pos.1'
VERSION : 0.1


VAR_TEMP
  TIMER_RESET : BOOL ;
  MAIN_SERVICE_1_SW : BOOL ;
  CONV_0_SERVICE_FWD : BOOL ;
  CONV_0_SERVICE_REV : BOOL ;
  RESET_1 : BOOL ;
  RESET_2 : BOOL ;
  PUSHER_PUSH : BOOL ;
END_VAR
BEGIN
NETWORK
TITLE =Conveyor 0 - Service

      A     "HMI_DB".ALL_SERVICE_ENABLE_SW;
      A     "HMI_DB".CONVEYOR_0_SERVICE_SW;
      A     "HMI_DB".SERVICE_SW_1_STATUS;
      =     #MAIN_SERVICE_1_SW;
//;
      A     #MAIN_SERVICE_1_SW;
      O     "M 14.0";
      JNB   PUS0;
      A     "HMI_DB".HMI_ROLLER_TEST_FWD_SSW;
      FP    "FP 168.3";
      R     "HMI_DB".HMI_ROLLER_TEST_REV_SSW;
      =     #RESET_1;
//;
      A     "HMI_DB".HMI_ROLLER_TEST_REV_SSW;
      FP    "FP 168.4";
      R     "HMI_DB".HMI_ROLLER_TEST_FWD_SSW;
      =     #RESET_2;
//;
      A(    ;
      O     #RESET_1;
      O     #RESET_2;
      )     ;
      L     S5T#1S;
      SF    "Timer 110";
//;
      A     "HMI_DB".HMI_ROLLER_TEST_FWD_SSW;
      AN    "Timer 110";
      =     #CONV_0_SERVICE_FWD;
//;
      A     "HMI_DB".HMI_ROLLER_TEST_REV_SSW;
      AN    "Timer 110";
      =     #CONV_0_SERVICE_REV;
//;
      A     "HMI_DB".HMI_PUSHER_0_TEST_SSW;
      =     #PUSHER_PUSH;
//;
      AN    #MAIN_SERVICE_1_SW;
      R     "HMI_DB".HMI_ROLLER_TEST_FWD_SSW;
      R     "HMI_DB".HMI_ROLLER_TEST_REV_SSW;

PUS0: R     #CONV_0_SERVICE_FWD;
      R     #CONV_0_SERVICE_REV;
      R     #RESET_1;
      R     #RESET_2;
      R     #PUSHER_PUSH;
      FP    "FP 158.0";
      =     "M 14.0";
NETWORK
TITLE =Function Keys <F5 > on HMI - Reset
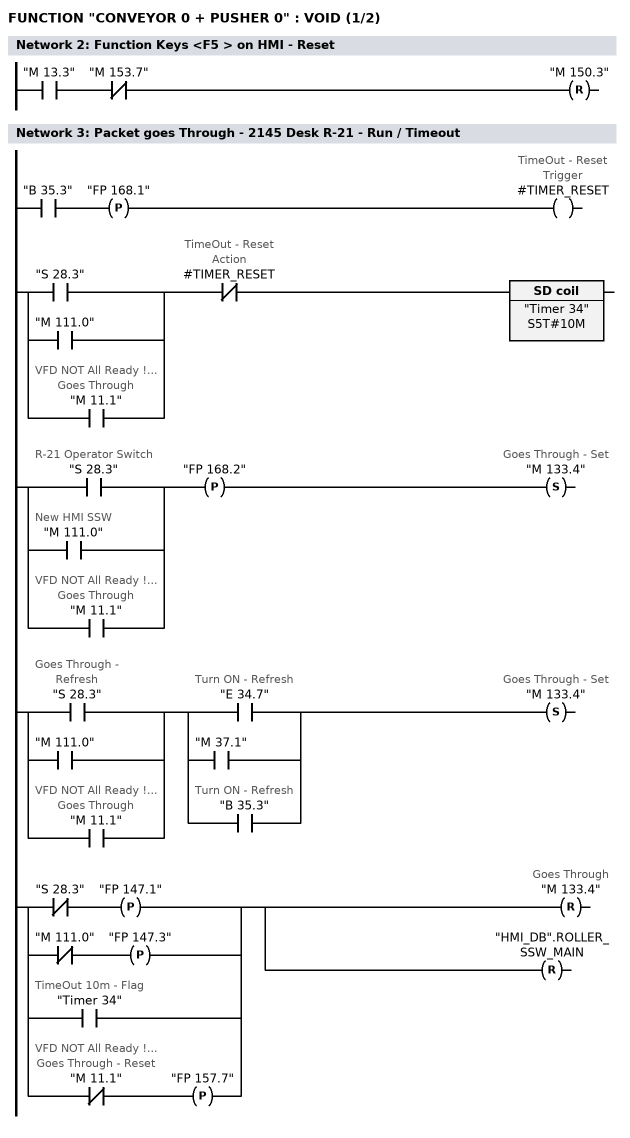

      A     "M 13.3";
      AN    "M 153.7";
      R     "M 150.3";
NETWORK
TITLE =Packet goes Through - 2145 Desk R-21 - Run / Timeout

      A     "B 35.3";
      FP    "FP 168.1";
      =     #TIMER_RESET; // TimeOut - Reset Trigger
//;
      A     "S 28.3";
      O     "M 111.0";
      O     "M 11.1"; // VFD NOT All Ready !... Goes Through
      AN    #TIMER_RESET; // TimeOut - Reset Action
      L     S5T#10M;
      SD    "Timer 34"; // TimeOut 10m
//;
      A     "S 28.3"; // R-21 Operator Switch
      O     "M 111.0"; // New HMI SSW
      O     "M 11.1"; // VFD NOT All Ready !... Goes Through
      FP    "FP 168.2"; // Turn ON - Pulse
      S     "M 133.4"; // Goes Through - Set
//;
      A     "S 28.3"; // Goes Through - Refresh
      O     "M 111.0";
      O     "M 11.1"; // VFD NOT All Ready !... Goes Through
      A(    ;
      O     "E 34.7"; // Turn ON - Refresh
      O     "M 37.1";
      O     "B 35.3"; // Turn ON - Refresh
      )     ;
      S     "M 133.4"; // Goes Through - Set
//;
      A(    ;
      O(    ;
      AN    "S 28.3";
      FP    "FP 147.1"; // Turn OFF - Pulse
      )     ;
      O(    ;
      AN    "M 111.0";
      FP    "FP 147.3"; // Turn OFF - Pulse
      O     "Timer 34"; // TimeOut 10m - Flag
      )     ;
      O(    ;
      AN    "M 11.1"; // VFD NOT All Ready !... Goes Through - Reset
      FP    "FP 157.7";
      )     ;
      )     ;
      R     "M 133.4"; // Goes Through
      R     "HMI_DB".ROLLER_SSW_MAIN;
NETWORK
TITLE =
//
//      A     "E 2.4"
//      S     "M 33.0"                    // Solid Detected ?
////;
//      A     "M 33.0"                    // Delay Timer - Start
//      L     S5T#300MS
//      SD    "Timer 26"                  // Debouncer 300mS
////;
//      A     "Timer 26"                  // Delayed Test Pulse
//      AN    "E 2.4"                     // Foul Detection
//      R     "M 33.0"                    // Not Detected !
////;
//      A     "Timer 26"                  // Delayed Test Pulse
//      A     "M 33.0"                    // Detection Comfirm !
//      =     "M 33.1"                    // Packet Height OK
//      R     "M 33.0"                    // Reset
//


NETWORK
TITLE =Packet Height - Sensing / Debouncing
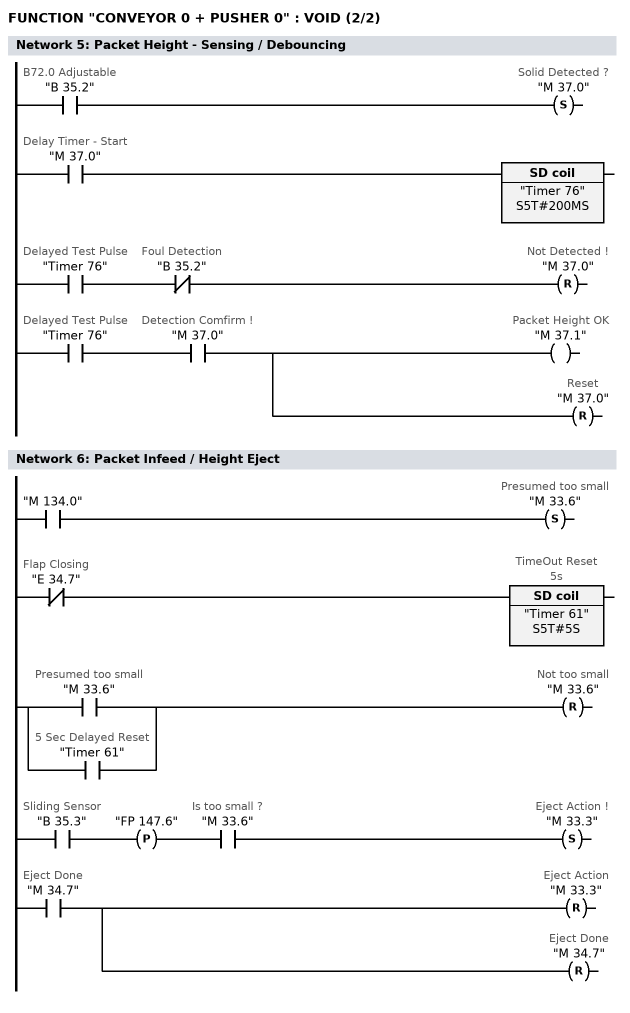

      A     "B 35.2"; // B72.0 Adjustable
      S     "M 37.0"; // Solid Detected ?
//;
      A     "M 37.0"; // Delay Timer - Start
      L     S5T#200MS;
      SD    "Timer 76"; // Debouncer 300mS
//;
      A     "Timer 76"; // Delayed Test Pulse
      AN    "B 35.2"; // Foul Detection
      R     "M 37.0"; // Not Detected !
//;
      A     "Timer 76"; // Delayed Test Pulse
      A     "M 37.0"; // Detection Comfirm !
      =     "M 37.1"; // Packet Height OK
      R     "M 37.0"; // Reset
NETWORK
TITLE =Packet Infeed / Height Eject

      A     "M 134.0";
      S     "M 33.6"; // Presumed too small
//;
      AN    "E 34.7"; // Flap Closing
      L     S5T#5S; // TimeOut Reset 5s
      SD    "Timer 61";
//;
      A     "M 33.6"; // Presumed too small
//    A     "M 33.1"                    // Packet Height OK ?
      O     "Timer 61"; // 5 Sec Delayed Reset
      R     "M 33.6"; // Not too small
//;
      A     "B 35.3"; // Sliding Sensor
      FP    "FP 147.6";
      A     "M 33.6"; // Is too small ?
      S     "M 33.3"; // Eject Action !
//;
      A     "M 34.7"; // Eject Done
      R     "M 33.3"; // Eject Action
      R     "M 34.7"; // Eject Done
NETWORK
TITLE =Eject Comfirmation

      A     "M 13.0";
      JNB   OUT1;

      A     "B 35.3";
      AN    "M 132.6"; // Not Triggered by Pusher
      S     "M 34.3"; // Eject Step 1
//;
      A     "B 35.4";
      AN    "M 132.6"; // Not Triggered by Pusher
      S     "M 34.4"; // Eject Step 2
//;
      A     "K 62.0"; // Conveyor 0 - Running
      A     "M 153.7";
      A     "M 34.3"; // Eject Step 1
      A     "M 34.4"; // Eject Step 2
      S     "M 34.5"; // Eject Step 3
//;
      A     "M 34.5"; // Eject Step 3
      AN    "B 35.4"; // Eject Step 4
      S     "M 34.7"; // Eject Done
      R     "M 34.3"; // Eject Step 1 - Reset
      R     "M 34.4"; // Eject Step 2 - Reset
      R     "M 34.5"; // Eject Step 3 - Reset
      R     "M 33.3"; // Eject Action - Reset
//;
      A     "M 132.5"; // Reset with Pusher Extend
      A     "B 35.4";
      R     "M 34.3"; // Eject Step 1 - Reset
      R     "M 34.4"; // Eject Step 2 - Reset
      R     "M 34.5"; // Eject Step 3 - Reset
      R     "M 33.3"; // Eject Action - Reset

OUT1: CLR   ;
NETWORK
TITLE =Packet goes Through - Conveyor 0 Man Run - LAUER F5
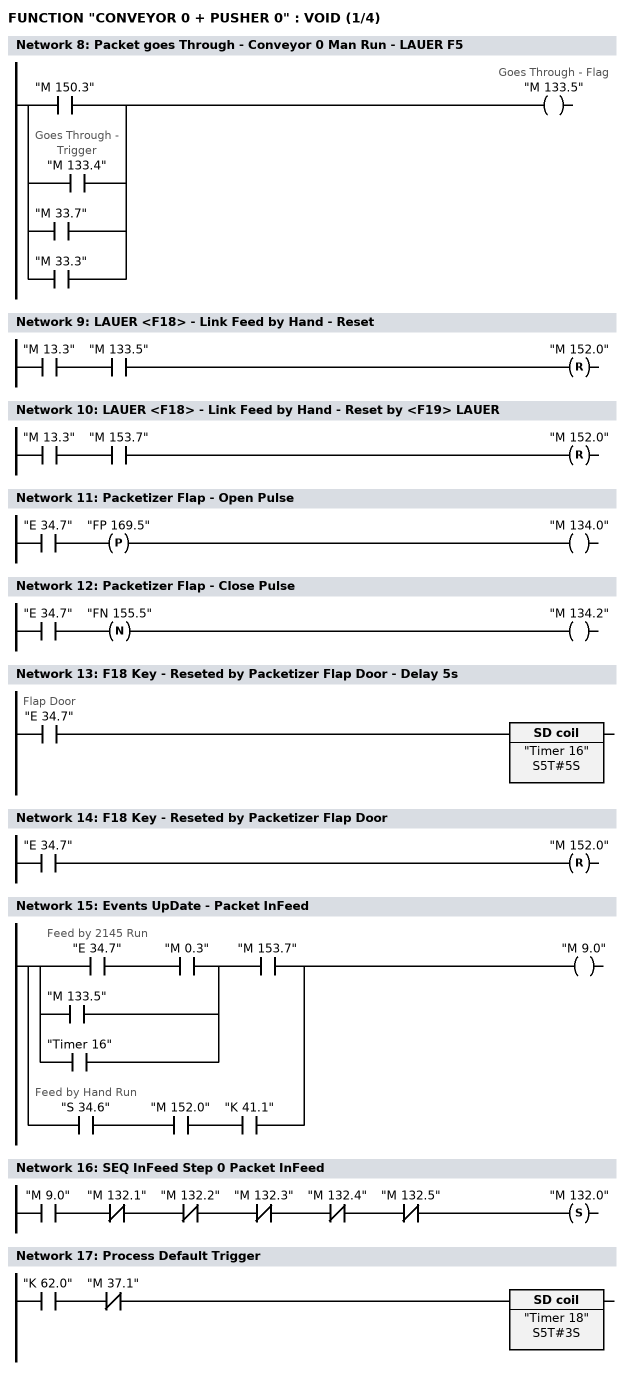

      O     "M 150.3";
      O     "M 133.4"; // Goes Through - Trigger
      O     "M 33.7";
      O     "M 33.3";
      =     "M 133.5"; // Goes Through - Flag
NETWORK
TITLE =LAUER <F18> - Link Feed by Hand - Reset

      A     "M 13.3";
      A     "M 133.5";
      R     "M 152.0";
NETWORK
TITLE =LAUER <F18> - Link Feed by Hand - Reset by <F19> LAUER

      A     "M 13.3";
      A     "M 153.7";
      R     "M 152.0";
NETWORK
TITLE =Packetizer Flap - Open Pulse

      A     "E 34.7";
      FP    "FP 169.5";
      =     "M 134.0";
NETWORK
TITLE =Packetizer Flap - Close Pulse

      A     "E 34.7";
      FN    "FN 155.5";
      =     "M 134.2";
NETWORK
TITLE =F18 Key - Reseted by Packetizer Flap Door - Delay 5s

      A     "E 34.7"; // Flap Door
      L     S5T#5S;
      SD    "Timer 16"; // Setup Mode Trigger
NETWORK
TITLE =F18 Key - Reseted by Packetizer Flap Door

      A     "E 34.7";
      R     "M 152.0";
NETWORK
TITLE =Events UpDate - Packet InFeed

      A(    ;
      A     "E 34.7"; // Feed by 2145 Run
      A     "M 0.3";
      O     "M 133.5";
      O     "Timer 16";
      A     "M 153.7";
      O     ;
      A     "S 34.6"; // Feed by Hand Run
      A     "M 152.0";
      A     "K 41.1";
      )     ;
      =     "M 9.0";
NETWORK
TITLE =SEQ InFeed Step 0 Packet InFeed

      A     "M 9.0";
      AN    "M 132.1";
      AN    "M 132.2";
      AN    "M 132.3";
      AN    "M 132.4";
      AN    "M 132.5";
      S     "M 132.0";
NETWORK
TITLE =Process Default Trigger

      A     "K 62.0";
      AN    "M 37.1";
      L     S5T#3S;
      SD    "Timer 18";
NETWORK
TITLE =Events UpDate
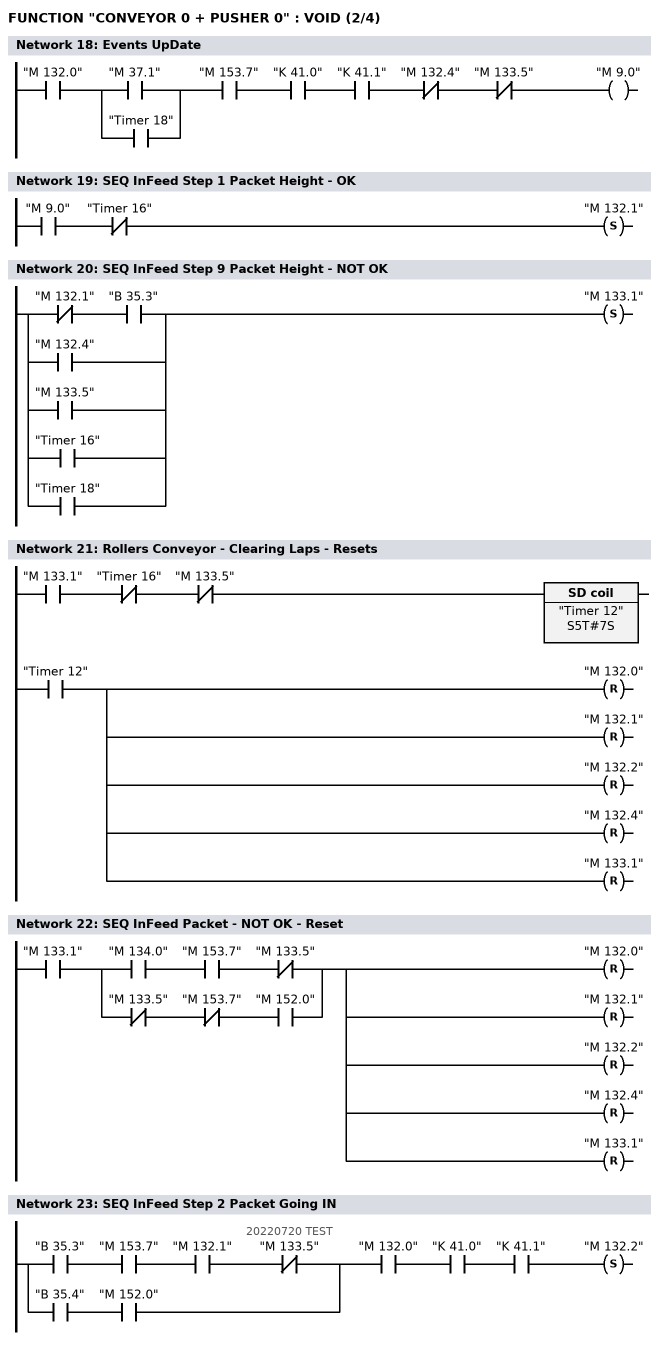

      A     "M 132.0";
      A(    ;
      O     "M 37.1";
      O     "Timer 18";
      )     ;
      A     "M 153.7";
      A     "K 41.0";
      A     "K 41.1";
      AN    "M 132.4";
      AN    "M 133.5";
      =     "M 9.0";
NETWORK
TITLE =SEQ InFeed Step 1 Packet Height - OK

      A     "M 9.0";
      AN    "Timer 16";
      S     "M 132.1";
NETWORK
TITLE =SEQ InFeed Step 9 Packet Height - NOT OK

      AN    "M 132.1";
      A     "B 35.3";
      O     "M 132.4";
      O     "M 133.5";
      O     "Timer 16";
      O     "Timer 18";
      S     "M 133.1";
NETWORK
TITLE =Rollers Conveyor - Clearing Laps - Resets

      A     "M 133.1";
      AN    "Timer 16";
      AN    "M 133.5";
      L     S5T#7S;
      SD    "Timer 12";
//;
      A     "Timer 12";
      R     "M 132.0";
      R     "M 132.1";
      R     "M 132.2";
      R     "M 132.4";
      R     "M 133.1";
NETWORK
TITLE =SEQ InFeed Packet - NOT OK - Reset

      A     "M 133.1";
      A(    ;
      A     "M 134.0";
      A     "M 153.7";
      AN    "M 133.5";
      O     ;
      AN    "M 133.5";
      AN    "M 153.7";
      A     "M 152.0";
      )     ;
      R     "M 132.0";
      R     "M 132.1";
      R     "M 132.2";
      R     "M 132.4";
      R     "M 133.1";
NETWORK
TITLE =SEQ InFeed Step 2 Packet Going IN

      A(    ;
      A     "B 35.3";
      A     "M 153.7";
      A     "M 132.1";
      AN    "M 133.5"; // 20220720 TEST
      O     ;
      A     "B 35.4";
      A     "M 152.0";
      )     ;
      A     "M 132.0";
      A     "K 41.0";
      A     "K 41.1";
      S     "M 132.2";
NETWORK
TITLE =SEQ InFeed Step 3 Conveyor Stop
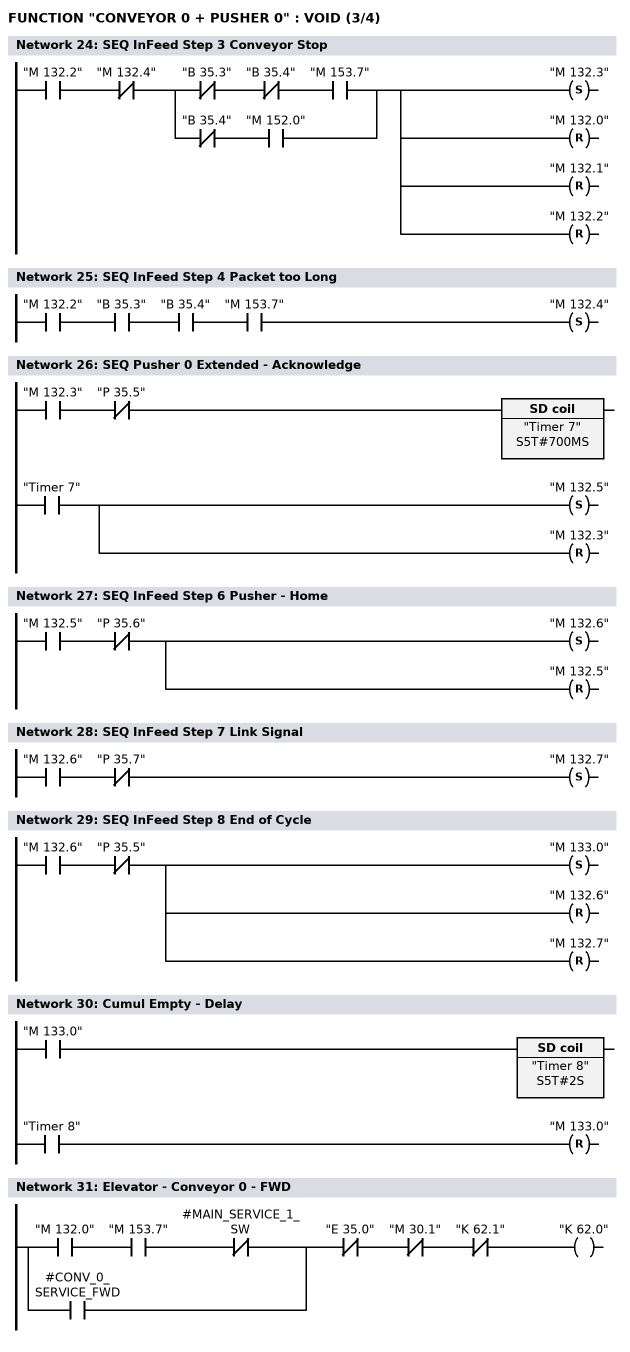

      A     "M 132.2";
      AN    "M 132.4";
      A(    ;
      AN    "B 35.3";
      AN    "B 35.4";
      A     "M 153.7";
      O     ;
      AN    "B 35.4";
      A     "M 152.0";
      )     ;
      S     "M 132.3";
      R     "M 132.0";
      R     "M 132.1";
      R     "M 132.2";
NETWORK
TITLE =SEQ InFeed Step 4 Packet too Long

      A     "M 132.2";
      A     "B 35.3";
      A     "B 35.4";
      A     "M 153.7";
      S     "M 132.4";
NETWORK
TITLE =SEQ Pusher 0 Extended - Acknowledge

      A     "M 132.3";
      AN    "P 35.5";
      L     S5T#700MS;
      SD    "Timer 7";
//;
      A     "Timer 7";
      S     "M 132.5";
      R     "M 132.3";
NETWORK
TITLE =SEQ InFeed Step 6 Pusher - Home

      A     "M 132.5";
      AN    "P 35.6";
      S     "M 132.6";
      R     "M 132.5";
NETWORK
TITLE =SEQ InFeed Step 7 Link Signal

      A     "M 132.6";
      AN    "P 35.7";
      S     "M 132.7";
NETWORK
TITLE =SEQ InFeed Step 8 End of Cycle

      A     "M 132.6";
      AN    "P 35.5";
      S     "M 133.0";
      R     "M 132.6";
      R     "M 132.7";
NETWORK
TITLE =Cumul Empty - Delay

      A     "M 133.0";
      L     S5T#2S;
      SD    "Timer 8";
//;
      A     "Timer 8";
      R     "M 133.0";
NETWORK
TITLE =Elevator - Conveyor 0 - FWD

      A(    ;
      A     "M 132.0";
      A     "M 153.7";
      AN    #MAIN_SERVICE_1_SW;
      O     #CONV_0_SERVICE_FWD;
      )     ;
      AN    "E 35.0";
      AN    "M 30.1";
      AN    "K 62.1";
      =     "K 62.0";
NETWORK
TITLE =Elevator - Conveyor 0 - REV
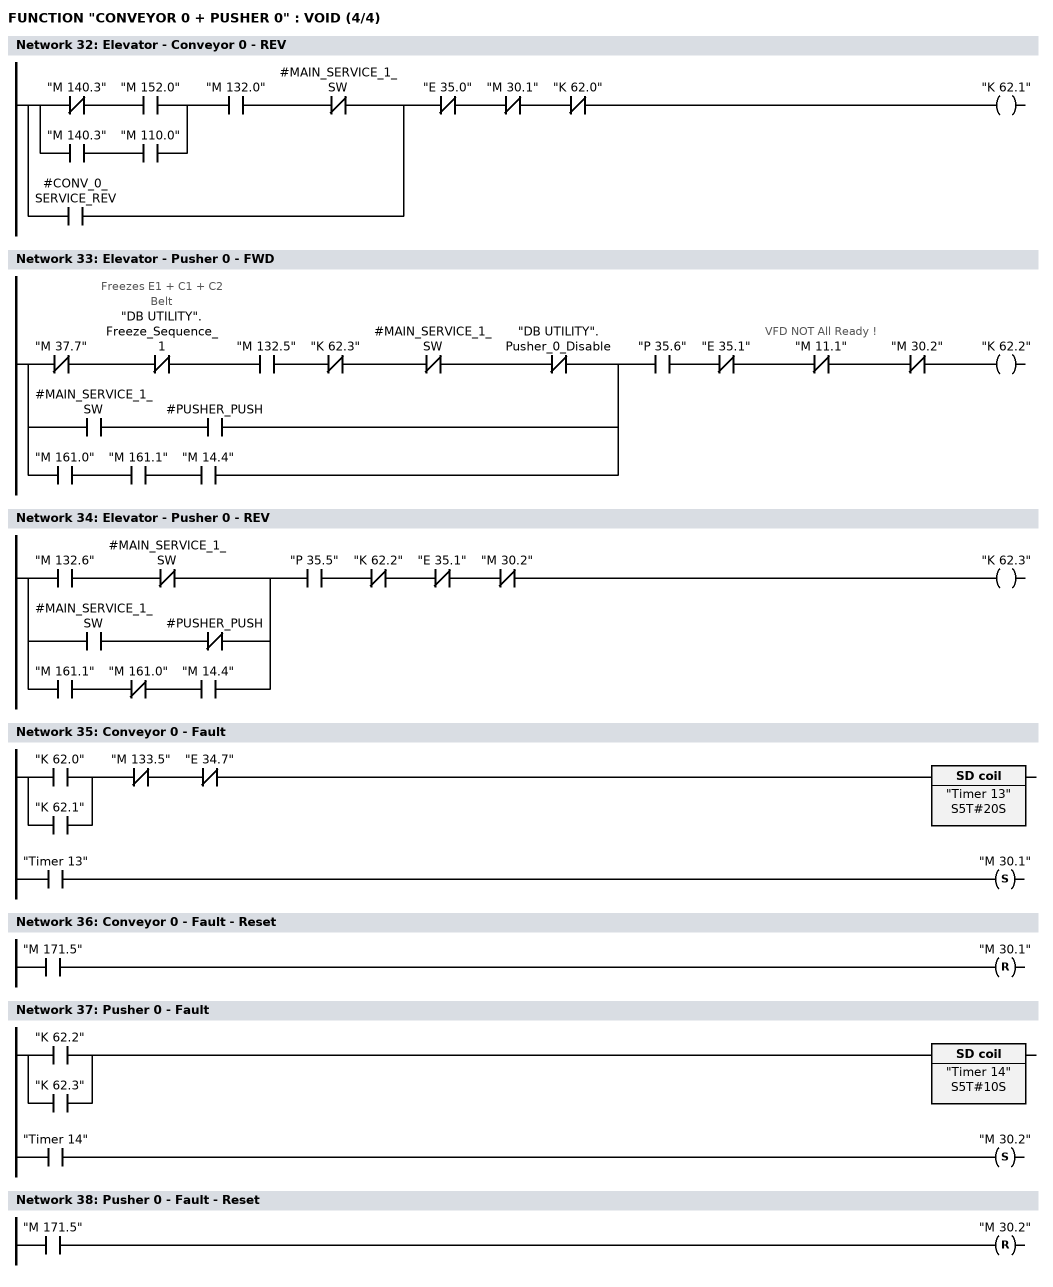

      A(    ;
      A(    ;
      AN    "M 140.3";
      A     "M 152.0";
      O     ;
      A     "M 140.3";
      A     "M 110.0";
      )     ;
      A     "M 132.0";
//     A     "M 152.0"
      AN    #MAIN_SERVICE_1_SW;
      O     #CONV_0_SERVICE_REV;
      )     ;
      AN    "E 35.0";
      AN    "M 30.1";
      AN    "K 62.0";
      =     "K 62.1";
NETWORK
TITLE =Elevator - Pusher 0 - FWD

      A(    ;
      AN    "M 37.7";
      AN    "DB UTILITY".Freeze_Sequence_1; //  Freezes E1 + C1 + C2 Belt
      A     "M 132.5";
      AN    "K 62.3";
      AN    #MAIN_SERVICE_1_SW;
      AN    "DB UTILITY".Pusher_0_Disable;
      O(    ;
      A     #MAIN_SERVICE_1_SW;
      A     #PUSHER_PUSH;
      )     ;
      O     ;
      A     "M 161.0";
      A     "M 161.1";
      A     "M 14.4";
      )     ;
      A     "P 35.6";
      AN    "E 35.1";
      AN    "M 11.1"; // VFD NOT All Ready !
      AN    "M 30.2";
      =     "K 62.2";
NETWORK
TITLE =Elevator - Pusher 0 - REV

      A(    ;
      A     "M 132.6";
      AN    #MAIN_SERVICE_1_SW;
      O(    ;
      A     #MAIN_SERVICE_1_SW;
      AN    #PUSHER_PUSH;
      )     ;
      O     ;
      A     "M 161.1";
      AN    "M 161.0";
      A     "M 14.4";
      )     ;
      A     "P 35.5";
      AN    "K 62.2";
      AN    "E 35.1";
      AN    "M 30.2";
      =     "K 62.3";
NETWORK
TITLE =Conveyor 0 - Fault

      A(    ;
      O     "K 62.0";
      O     "K 62.1";
      )     ;
      AN    "M 133.5";
      AN    "E 34.7";
      L     S5T#20S;
      SD    "Timer 13";
//;
      A     "Timer 13";
      S     "M 30.1";
NETWORK
TITLE =Conveyor 0 - Fault - Reset

      A     "M 171.5";
      R     "M 30.1";
NETWORK
TITLE =Pusher 0 - Fault

      A(    ;
      O     "K 62.2";
      O     "K 62.3";
      )     ;
      L     S5T#10S;
      SD    "Timer 14";
//;
      A     "Timer 14";
      S     "M 30.2";
NETWORK
TITLE =Pusher 0 - Fault - Reset

      A     "M 171.5";
      R     "M 30.2";
END_FUNCTION

FUNCTION "ELEVATOR + PUSHER 1" : VOID
TITLE =Elevator + Pusher 1   Pos.2  FC1016
//
NAME : POS_2
VERSION : 0.0


VAR_TEMP
  ELEVATOR_UP_OUT : BOOL ;
  ELEVATOR_DN_OUT : BOOL ;
  MAIN_SERVICE_1_SW : BOOL ;
  ELEVATOR_SERVICE_SW : BOOL ;
  ELEVATOR_DN_PB : BOOL ;
  ELEVATOR_UP_PB : BOOL ;
  ELEVATOR_ROUNDTRIP : BOOL ;
  PUSHER_PUSH : BOOL ;
  INITIALISATION : BOOL ;
  BRAKE_RELEASE_OK : BOOL ;
  BRAKE_CONTACTOR_KO : BOOL ;
END_VAR
BEGIN
NETWORK
TITLE =Elevator - Health OK
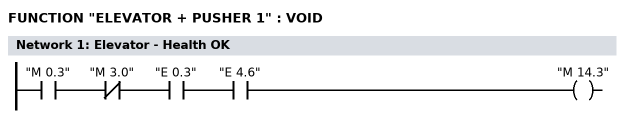

      A     "M 0.3";
      AN    "M 3.0";
      A     "E 0.3";
      A     "E 4.6";
      =     "M 14.3";
NETWORK
TITLE =Elevator - Service

      A     "HMI_DB".ALL_SERVICE_ENABLE_SW;
      A     "HMI_DB".ELEVATOR_SERVICE_SW;
      A     "HMI_DB".SERVICE_SW_1_STATUS;
      =     #MAIN_SERVICE_1_SW;
//;
      A     #MAIN_SERVICE_1_SW;
      O     "M 14.1";
      JNB   PUS1;
      A     "HMI_DB".HMI_ELEVATOR_SERVICE_SSW;
      =     #ELEVATOR_SERVICE_SW;
      S     "DB UTILITY".Pusher_0_Disable;
//;
      A     #ELEVATOR_SERVICE_SW;
      A(    ;
      A     "HMI_DB".HMI_ELEVATOR_TEST_DN_SSW;
      )     ;
      =     #ELEVATOR_DN_PB;
//;
      A     #ELEVATOR_SERVICE_SW;
      A(    ;
      A     "HMI_DB".HMI_ELEVATOR_TEST_UP_SSW;
      )     ;
      =     #ELEVATOR_UP_PB;
//;
      A     #MAIN_SERVICE_1_SW;
      AN    #ELEVATOR_SERVICE_SW;
      A     "HMI_DB".ELEVATOR_ROUND_TRIP_SSW;
      =     #ELEVATOR_ROUNDTRIP;
//;
      A     "HMI_DB".HMI_PUSHER_1_TEST_SSW;
      =     #PUSHER_PUSH;
//;
      AN    #MAIN_SERVICE_1_SW;
      R     "HMI_DB".HMI_ELEVATOR_SERVICE_SSW;
      R     "HMI_DB".HMI_ELEVATOR_TEST_DN_SSW;
      R     "HMI_DB".HMI_ELEVATOR_TEST_UP_SSW;
      R     "DB UTILITY".Pusher_0_Disable;

PUS1: R     #ELEVATOR_SERVICE_SW;
      R     #ELEVATOR_DN_PB;
      R     #ELEVATOR_UP_PB;
      R     #ELEVATOR_ROUNDTRIP;
      R     #PUSHER_PUSH;
      FP    "FP 158.1";
      =     "M 14.1";
//;
      A     "HMI_DB".SERVICE_INIT_PB;
      A     #ELEVATOR_SERVICE_SW;
      A     #MAIN_SERVICE_1_SW;
      =     #INITIALISATION;
NETWORK
TITLE =Elevator - Manual Run - Conditions
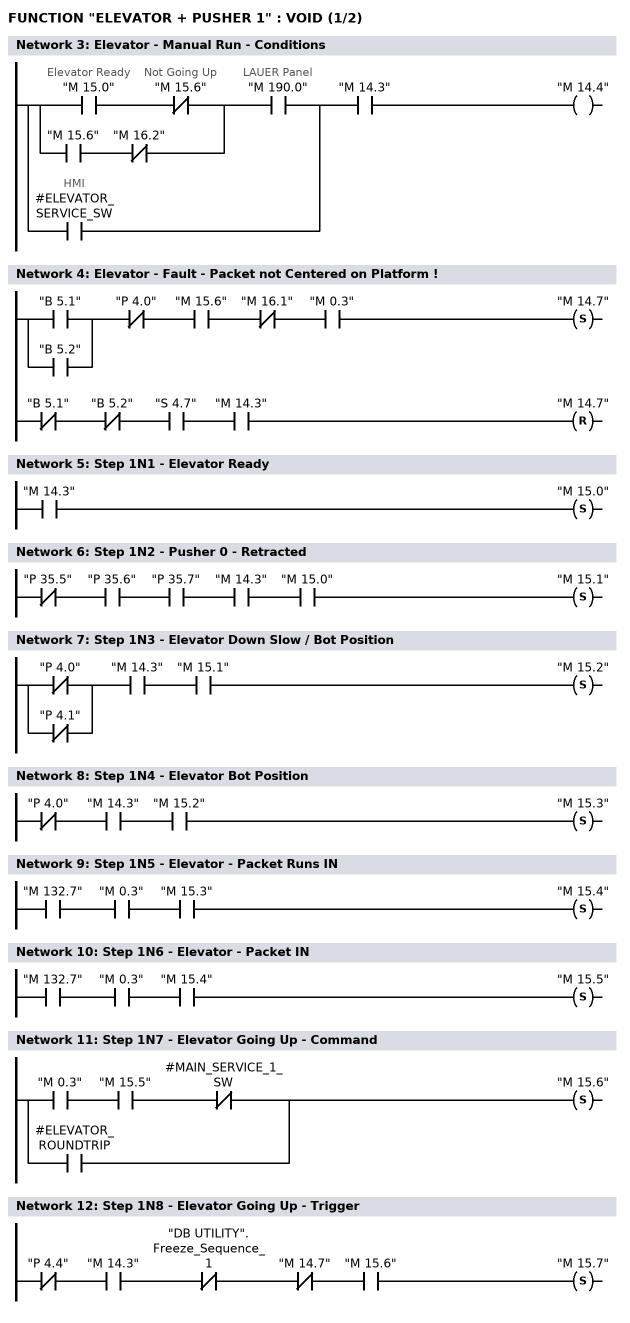

      A(    ;
      A     "M 15.0"; // Elevator Ready
      AN    "M 15.6"; // Not Going Up
      O     ; // or
      A     "M 15.6";
      AN    "M 16.2";
      )     ;
      A     "M 190.0"; // LAUER Panel
      O     #ELEVATOR_SERVICE_SW; // HMI
      A     "M 14.3";
      =     "M 14.4";
NETWORK
TITLE =Elevator - Fault - Packet not Centered on Platform !

      A(    ;
      O     "B 5.1";
      O     "B 5.2";
      )     ;
      AN    "P 4.0";
      A     "M 15.6";
      AN    "M 16.1";
      A     "M 0.3";
      S     "M 14.7";
//;
      AN    "B 5.1";
      AN    "B 5.2";
      A     "S 4.7";
      A     "M 14.3";
      R     "M 14.7";
NETWORK
TITLE =Step 1N1 - Elevator Ready

      A     "M 14.3";
      S     "M 15.0";
NETWORK
TITLE =Step 1N2 - Pusher 0 - Retracted

      AN    "P 35.5";
      A     "P 35.6";
      A     "P 35.7";
      A     "M 14.3";
      A     "M 15.0";
      S     "M 15.1";
NETWORK
TITLE =Step 1N3 - Elevator Down Slow / Bot Position

      A(    ;
      ON    "P 4.0";
      ON    "P 4.1";
      )     ;
      A     "M 14.3";
      A     "M 15.1";
      S     "M 15.2";
NETWORK
TITLE =Step 1N4 - Elevator Bot Position

      AN    "P 4.0";
      A     "M 14.3";
      A     "M 15.2";
      S     "M 15.3";
NETWORK
TITLE =Step 1N5 - Elevator - Packet Runs IN

      A     "M 132.7";
      A     "M 0.3";
      A     "M 15.3";
      S     "M 15.4";
NETWORK
TITLE =Step 1N6 - Elevator - Packet IN

      A     "M 132.7";
      A     "M 0.3";
      A     "M 15.4";
      S     "M 15.5";
NETWORK
TITLE =Step 1N7 - Elevator Going Up - Command

      A     "M 0.3";
      A     "M 15.5";
      AN    #MAIN_SERVICE_1_SW;
      O     #ELEVATOR_ROUNDTRIP;
      S     "M 15.6";
NETWORK
TITLE =Step 1N8 - Elevator Going Up - Trigger

      AN    "P 4.4";
      A     "M 14.3";
      AN    "DB UTILITY".Freeze_Sequence_1;
      AN    "M 14.7";
      A     "M 15.6";
      S     "M 15.7";
NETWORK
TITLE =Step 1N9 - Elevator Going Up - Slow
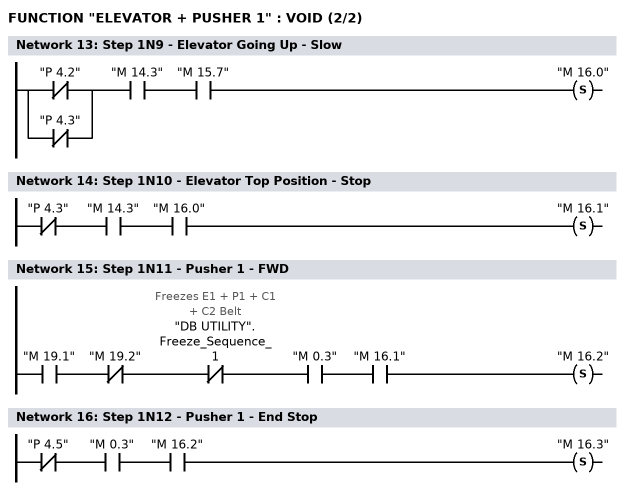

      A(    ;
      ON    "P 4.2";
      ON    "P 4.3";
      )     ;
      A     "M 14.3";
      A     "M 15.7";
      S     "M 16.0";
NETWORK
TITLE =Step 1N10 - Elevator Top Position - Stop

      AN    "P 4.3";
      A     "M 14.3";
      A     "M 16.0";
      S     "M 16.1";
NETWORK
TITLE =Step 1N11 - Pusher 1 - FWD

      A     "M 19.1";
      AN    "M 19.2";
      AN    "DB UTILITY".Freeze_Sequence_1; //  Freezes E1 + P1 + C1 + C2 Belt
      A     "M 0.3";
      A     "M 16.1";
      S     "M 16.2";
NETWORK
TITLE =Step 1N12 - Pusher 1 - End Stop

      AN    "P 4.5";
      A     "M 0.3";
      A     "M 16.2";
      S     "M 16.3";
NETWORK
TITLE =Soft Timer 15 Reset

      A     "M 16.3";
      AN    "M 16.4";
      A     "M 14.3";
      A     "M 0.3";
      JCN   R151;
      JU    E151;

R151: L     L#0;
      T     "DB UTILITY".T15_ET;
      R     "DB UTILITY".T15_DN;

E151: NOP   0;

NETWORK
TITLE =Soft Timer 15 Add

      A     "M 16.3";
      AN    "M 16.4";
      A     "M 14.3";
      A     "M 0.3";
      AN    "DB UTILITY".Freeze_Sequence_1;
      AN    "DB UTILITY".T15_DN;
      JCN   E152;

      L     "DB UTILITY".T15_ET;
      L     "DB UTILITY".Scan_Cycle_Previous;
      ITD   ;
      +D    ;
      T     "DB UTILITY".T15_ET;

E152: NOP   0;

NETWORK
TITLE =Soft Timer 15 Done 100mS
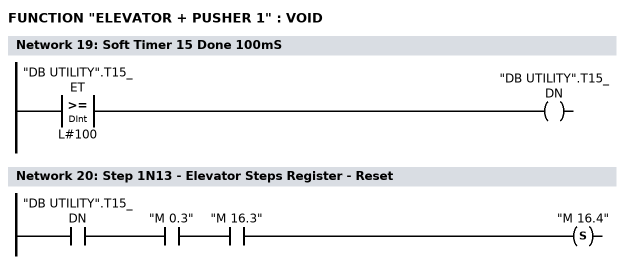

      L     "DB UTILITY".T15_ET;
      L     L#100;
      >=D   ;
      =     "DB UTILITY".T15_DN;

NETWORK
TITLE =Step 1N13 - Elevator Steps Register - Reset

      A     "DB UTILITY".T15_DN;
      A     "M 0.3";
      A     "M 16.3";
      S     "M 16.4";
NETWORK
TITLE =Elevator Steps Register - Reset

      A(    ;
      A     "M 190.0";
      A     "M 171.4";
      A     "M 171.5";
      O     "M 16.4";
      O     #INITIALISATION;
      O     "DB UTILITY".Elevator_Disable;
      )     ;
      A     "M 0.3";
      JC    M001;
      JU    M002;

M001: L     W#16#0;
      T     "MW 15";

M002: CLR   ;
NETWORK
TITLE =Trans System - Ready -> Tuber 2145
